FOR _bitIdx := 0 TO 15 DO
    IF (_reg.managedBitMask AND SHL(WORD#1, _bitIdx)) <> 0 THEN
        _sigIdx := _reg.arrSignalIndex[_bitIdx];

        IF _sigIdx > 0 THEN
            _pData := inpPtrWriteData + UINT_TO_DWORD(_sigIdx - 1) * SIZEOF(ST_MBWriteData);

            IF _pData^.valueBool THEN
                _baseValue := _baseValue OR SHL(WORD#1, _bitIdx);
            ELSE
                _baseValue := _baseValue AND NOT SHL(WORD#1, _bitIdx);
            END_IF
        END_IF
    END_IF
END_FOR

_reg.writeValue := _baseValue;
END_METHOD

METHOD PRIVATE checkReadComplete : BOOL
CASE _arrReadBlocks[_currentBlockIdx].functionCode OF
    1:
        fbMbReadCoils(bExecute := FALSE);
        checkReadComplete := NOT fbMbReadCoils.bBusy;
    2:
        fbMbReadInputs(bExecute := FALSE);
        checkReadComplete := NOT fbMbReadInputs.bBusy;
    3:
        fbMbReadRegs(bExecute := FALSE);
        checkReadComplete := NOT fbMbReadRegs.bBusy;
    4:
        fbMbReadInputRegs(bExecute := FALSE);
        checkReadComplete := NOT fbMbReadInputRegs.bBusy;
ELSE
    // RMW read path uses fbMbReadRegs unconditionally.
    fbMbReadRegs(bExecute := FALSE);
    checkReadComplete := NOT fbMbReadRegs.bBusy;
END_CASE
END_METHOD

METHOD PRIVATE checkStaleData
VAR
    _i          : UINT;
    _pResult    : POINTER TO ST_MBReadResult;
    _elapsed    : TIME;
END_VAR
_elapsed := TIME() - _lastGoodReadTime;

IF _elapsed > cfgStaleThreshold THEN
    FOR _i := 1 TO cfgReadSignalCount DO
        _pResult := inpPtrReadResults + UINT_TO_DWORD(_i - 1) * SIZEOF(ST_MBReadResult);

        IF _pResult^.quality = E_SignalQuality.Good THEN
            _pResult^.quality := E_SignalQuality.UncertainStale;
        END_IF
    END_FOR
END_IF
END_METHOD

METHOD PRIVATE checkWriteComplete : BOOL
IF _state = E_DriverState.WriteWait THEN
    IF _arrWriteBlocks[_currentBlockIdx].area = E_MBArea.Coils THEN
        fbMbWriteCoils(bExecute := FALSE);
        checkWriteComplete := NOT fbMbWriteCoils.bBusy;
    ELSE
        fbMbWriteRegs(bExecute := FALSE);
        checkWriteComplete := NOT fbMbWriteRegs.bBusy;
    END_IF
ELSE
    fbMbWriteSingleReg(bExecute := FALSE);
    checkWriteComplete := NOT fbMbWriteSingleReg.bBusy;
END_IF
END_METHOD

// Recover a Faulted (or errored) driver without toggling inpEnable: it restarts from Init on
// the next cycle() — re-parses the configuration and resumes polling. No effect while disabled.
METHOD PUBLIC cmdReset : BOOL
IF inpEnable THEN
    _state := E_DriverState.Init;
    _resetRequest := TRUE;
    cmdReset := TRUE;
END_IF
END_METHOD

METHOD PRIVATE combineWords : DWORD
VAR_INPUT
    inpWord0        : WORD;
    inpWord1        : WORD;
END_VAR
IF cfgWordOrder = E_WordOrder.BigEndian THEN
    combineWords := SHL(WORD_TO_DWORD(inpWord0), 16) OR WORD_TO_DWORD(inpWord1);
ELSE
    combineWords := SHL(WORD_TO_DWORD(inpWord1), 16) OR WORD_TO_DWORD(inpWord0);
END_IF
END_METHOD

PROPERTY PUBLIC commandDelay : TIME
GET
commandDelay := cfgCommandDelay;
END_GET
SET
IF NOT _initialized THEN
    cfgCommandDelay := commandDelay;
END_IF
END_SET
END_PROPERTY

METHOD PUBLIC cycle
VAR
    _risingEnable   : BOOL;
END_VAR
_risingEnable := inpEnable AND NOT _enablePrev;
_enablePrev := inpEnable;

IF NOT inpEnable THEN
    disable();
    RETURN;
END_IF

IF _initialized AND _socketConnected THEN
    stsStatus.timeSinceLastGoodRead := TIME() - _lastGoodReadTime;
    stsStatus.timeSinceLastGoodWrite := TIME() - _lastGoodWriteTime;
END_IF

CASE _state OF

    E_DriverState.Init:
        IF _risingEnable OR _resetRequest THEN
            _resetRequest := FALSE;
            reset();
            _state := E_DriverState.ParseConfig;
        END_IF

    E_DriverState.ParseConfig:
        IF parseAllConfigs() THEN
            _state := E_DriverState.OptimizeBlocks;
        ELSE
            stsError := TRUE;
            _state := E_DriverState.Error;
        END_IF

    E_DriverState.OptimizeBlocks:
        optimizeReadBlocks();
        optimizeWriteBlocks();
        identifyBitRegisters();

        stsStatus.readBlockCount := _readBlockCount;
        stsStatus.writeBlockCount := _writeBlockCount;
        stsStatus.bitRegisterCount := _bitRegisterCount;

        _initialized := TRUE;
        _state := E_DriverState.Connecting;

    E_DriverState.Connecting:
        // Tc2_ModbusCaller manages TCP internally per FB call; no explicit connect.
        // Treat the driver as "ready to talk" once configs are parsed.
        _socketConnected := TRUE;
        _connectAttempts := 0;
        stsStatus.connected := TRUE;
        stsStatus.reconnectAttempts := 0;
        _lastGoodReadTime := TIME();
        _lastGoodWriteTime := TIME();
        _state := E_DriverState.Ready;

    E_DriverState.ConnectWait:
        // Vestigial state retained for E_DriverState compatibility; transition to Ready.
        _state := E_DriverState.Ready;

    E_DriverState.ReconnectWait:
        tonReconnectDelay(IN := TRUE, PT := cfgReconnectDelay);
        IF tonReconnectDelay.Q THEN
            tonReconnectDelay(IN := FALSE);
            _socketConnected := TRUE;
            stsStatus.connected := TRUE;
            _state := E_DriverState.Ready;
        END_IF

    E_DriverState.Disconnecting:
        // No socket to disconnect (Tc2_ModbusCaller is per-call).
        _socketConnected := FALSE;
        stsStatus.connected := FALSE;
        stsStatus.readCycleActive := FALSE;
        stsStatus.writeCycleActive := FALSE;
        _consecFailures := 0;           // the retry gets its own maxConsecFails budget
        _state := E_DriverState.DisconnectWait;

    E_DriverState.DisconnectWait:
        IF _disconnectPending THEN
            _disconnectPending := FALSE;
            tonReconnectDelay(IN := FALSE);
            _state := E_DriverState.ReconnectWait;
        ELSE
            _state := E_DriverState.Init;
        END_IF

    E_DriverState.Ready:
        tonPollInterval(IN := TRUE, PT := cfgPollInterval);
        IF tonPollInterval.Q THEN
            tonPollInterval(IN := FALSE);
            IF _readBlockCount > 0 THEN
                _state := E_DriverState.ReadStart;
                RETURN;
            END_IF
        END_IF

        tonWriteInterval(IN := TRUE, PT := cfgWriteCycleInterval);
        IF tonWriteInterval.Q THEN
            tonWriteInterval(IN := FALSE);
            IF NOT inpHoldWrites AND (_writeBlockCount > 0 OR _bitRegisterCount > 0) THEN
                _state := E_DriverState.WriteStart;
                RETURN;
            END_IF
        END_IF

        checkStaleData();

    E_DriverState.ReadStart:
        _currentBlockIdx := 1;
        _readCycleFailed := FALSE;
        stsStatus.readCycleActive := TRUE;
        _state := E_DriverState.ReadSend;

    E_DriverState.ReadSend:
        IF _currentBlockIdx > _readBlockCount THEN
            _state := E_DriverState.ReadComplete;
        ELSE
            sendReadRequest(_currentBlockIdx);
            _state := E_DriverState.ReadWait;
        END_IF

    E_DriverState.ReadWait:
        tonTimeout(IN := TRUE, PT := cfgTimeout);

        IF checkReadComplete() THEN
            tonTimeout(IN := FALSE);
            IF readSucceeded() THEN
                processReadBlock(_currentBlockIdx);
                _consecFailures := 0;
            ELSE
                handleBlockError(_currentBlockIdx, TRUE);
            END_IF
            IF _state = E_DriverState.ReadWait THEN   // the error handler may have moved us to Disconnecting/Faulted
                _state := E_DriverState.ReadDelay;
            END_IF

        ELSIF tonTimeout.Q THEN
            tonTimeout(IN := FALSE);
            handleBlockError(_currentBlockIdx, TRUE);
            IF _state = E_DriverState.ReadWait THEN   // the error handler may have moved us to Disconnecting/Faulted
                _state := E_DriverState.ReadDelay;
            END_IF
        END_IF

    E_DriverState.ReadDelay:
        tonCommandDelay(IN := TRUE, PT := cfgCommandDelay);
        IF tonCommandDelay.Q THEN
            tonCommandDelay(IN := FALSE);
            _currentBlockIdx := _currentBlockIdx + 1;
            _state := E_DriverState.ReadSend;
        END_IF

    E_DriverState.ReadComplete:
        stsStatus.readCycleActive := FALSE;
        stsStatus.totalReadCycles := stsStatus.totalReadCycles + 1;
        // Only a cycle in which EVERY block succeeded is a good read. Stamping it regardless
        // kept timeSinceLastGoodRead near zero (and stale marking off) while every read failed.
        IF NOT _readCycleFailed THEN
            _lastGoodReadTime := TIME();
            _connectAttempts := 0;      // link proven again: the reconnect budget starts over
            stsStatus.reconnectAttempts := 0;
        END_IF
        _state := E_DriverState.Ready;

    E_DriverState.WriteStart:
        _currentBlockIdx := 1;
        _writeCycleFailed := FALSE;
        _currentRmwIdx := 0;
        stsStatus.writeCycleActive := TRUE;
        _state := E_DriverState.WriteSend;

    E_DriverState.WriteSend:
        WHILE _currentBlockIdx <= _writeBlockCount DO
            IF NOT _arrWriteBlocks[_currentBlockIdx].containsBitSignals THEN
                packAndSendWriteBlock(_currentBlockIdx);
                _state := E_DriverState.WriteWait;
                RETURN;
            END_IF
            _currentBlockIdx := _currentBlockIdx + 1;
        END_WHILE

        IF _currentRmwIdx < _bitRegisterCount THEN
            _currentRmwIdx := _currentRmwIdx + 1;
            _state := E_DriverState.RmwReadSend;
        ELSE
            _state := E_DriverState.WriteComplete;
        END_IF

    E_DriverState.WriteWait:
        tonTimeout(IN := TRUE, PT := cfgTimeout);

        IF checkWriteComplete() THEN
            tonTimeout(IN := FALSE);
            IF writeSucceeded() THEN
                updateWriteStatus(_currentBlockIdx, TRUE);
                _consecFailures := 0;
            ELSE
                handleBlockError(_currentBlockIdx, FALSE);
                updateWriteStatus(_currentBlockIdx, FALSE);
            END_IF
            IF _state = E_DriverState.WriteWait THEN   // the error handler may have moved us to Disconnecting/Faulted
                _state := E_DriverState.WriteDelay;
            END_IF

        ELSIF tonTimeout.Q THEN
            tonTimeout(IN := FALSE);
            handleBlockError(_currentBlockIdx, FALSE);
            updateWriteStatus(_currentBlockIdx, FALSE);
            IF _state = E_DriverState.WriteWait THEN   // the error handler may have moved us to Disconnecting/Faulted
                _state := E_DriverState.WriteDelay;
            END_IF
        END_IF

    E_DriverState.WriteDelay:
        tonCommandDelay(IN := TRUE, PT := cfgCommandDelay);
        IF tonCommandDelay.Q THEN
            tonCommandDelay(IN := FALSE);
            _currentBlockIdx := _currentBlockIdx + 1;
            _state := E_DriverState.WriteSend;
        END_IF

    E_DriverState.RmwReadSend:
        sendRmwReadRequest(_currentRmwIdx);
        _state := E_DriverState.RmwReadWait;

    E_DriverState.RmwReadWait:
        tonTimeout(IN := TRUE, PT := cfgTimeout);

        IF checkReadComplete() THEN
            tonTimeout(IN := FALSE);
            IF readSucceeded() THEN
                _arrBitRegisters[_currentRmwIdx].readValue := _arrRawReadBuffer[0];
                _state := E_DriverState.RmwModify;
            ELSE
                handleRmwError(_currentRmwIdx);
                IF _state = E_DriverState.RmwReadWait THEN   // the error handler may have moved us to Disconnecting/Faulted
                    _state := E_DriverState.RmwDelay;
                END_IF
            END_IF

        ELSIF tonTimeout.Q THEN
            tonTimeout(IN := FALSE);
            handleRmwError(_currentRmwIdx);
            IF _state = E_DriverState.RmwReadWait THEN   // the error handler may have moved us to Disconnecting/Faulted
                _state := E_DriverState.RmwDelay;
            END_IF
        END_IF

    E_DriverState.RmwModify:
        applyBitModifications(_currentRmwIdx);
        _state := E_DriverState.RmwWriteSend;

    E_DriverState.RmwWriteSend:
        sendRmwWriteRequest(_currentRmwIdx);
        _state := E_DriverState.RmwWriteWait;

    E_DriverState.RmwWriteWait:
        tonTimeout(IN := TRUE, PT := cfgTimeout);

        IF checkWriteComplete() THEN
            tonTimeout(IN := FALSE);
            IF writeSucceeded() THEN
                updateRmwStatus(_currentRmwIdx, TRUE);
                _consecFailures := 0;
            ELSE
                handleRmwError(_currentRmwIdx);
                updateRmwStatus(_currentRmwIdx, FALSE);
            END_IF
            IF _state = E_DriverState.RmwWriteWait THEN   // the error handler may have moved us to Disconnecting/Faulted
                _state := E_DriverState.RmwDelay;
            END_IF

        ELSIF tonTimeout.Q THEN
            tonTimeout(IN := FALSE);
            handleRmwError(_currentRmwIdx);
            updateRmwStatus(_currentRmwIdx, FALSE);
            IF _state = E_DriverState.RmwWriteWait THEN   // the error handler may have moved us to Disconnecting/Faulted
                _state := E_DriverState.RmwDelay;
            END_IF
        END_IF

    E_DriverState.RmwDelay:
        tonCommandDelay(IN := TRUE, PT := cfgCommandDelay);
        IF tonCommandDelay.Q THEN
            tonCommandDelay(IN := FALSE);
            IF _currentRmwIdx < _bitRegisterCount THEN
                _currentRmwIdx := _currentRmwIdx + 1;
                _state := E_DriverState.RmwReadSend;
            ELSE
                _state := E_DriverState.WriteComplete;
            END_IF
        END_IF

    E_DriverState.WriteComplete:
        stsStatus.writeCycleActive := FALSE;
        stsStatus.totalWriteCycles := stsStatus.totalWriteCycles + 1;
        IF NOT _writeCycleFailed THEN
            _lastGoodWriteTime := TIME();
        END_IF
        _state := E_DriverState.Ready;

    E_DriverState.Error:
        stsError := TRUE;
        stsStatus.totalErrors := stsStatus.totalErrors + 1;
        _disconnectPending := TRUE;
        _state := E_DriverState.Disconnecting;

    E_DriverState.Faulted:
        stsStatus.faulted := TRUE;
        stsError := TRUE;

END_CASE

stsStatus.currentState := _state;
stsStatus.consecutiveFailures := _consecFailures;
END_METHOD

METHOD PRIVATE dintToWords
VAR_INPUT
    inpValue        : DINT;
END_VAR
VAR_OUTPUT
    stsWord0        : WORD;
    stsWord1        : WORD;
END_VAR
VAR
    _dword          : DWORD;
    _w0, _w1        : WORD;
END_VAR
_dword := DINT_TO_DWORD(inpValue);
splitDword(inpValue := _dword, stsWord0 => _w0, stsWord1 => _w1);
stsWord0 := swapBytes(_w0);
stsWord1 := swapBytes(_w1);
END_METHOD

METHOD PRIVATE disable
// Tc2_ModbusCaller has no socket to tear down explicitly.
_socketConnected := FALSE;

tonPollInterval(IN := FALSE);
tonWriteInterval(IN := FALSE);
tonCommandDelay(IN := FALSE);
tonTimeout(IN := FALSE);
tonReconnectDelay(IN := FALSE);

// Back to Init from ANY state, Faulted included: re-enabling restarts the driver. (Faulted used
// to survive a disable, which left a faulted driver dead until the PLC restarted.)
_state := E_DriverState.Init;
_resetRequest := FALSE;

_initialized := FALSE;
stsStatus.connected := FALSE;
stsStatus.readCycleActive := FALSE;
stsStatus.writeCycleActive := FALSE;
END_METHOD

METHOD PRIVATE handleBlockError
VAR_INPUT
    inpBlockIdx : UINT;
    inpIsRead   : BOOL;
END_VAR
VAR
    _block      : REFERENCE TO ST_ReadBlock;
    _i          : UINT;
    _sigIdx     : UINT;
    _pResult    : POINTER TO ST_MBReadResult;
END_VAR
_consecFailures := _consecFailures + 1;
stsStatus.totalErrors := stsStatus.totalErrors + 1;
IF inpIsRead THEN
    _readCycleFailed := TRUE;
ELSE
    _writeCycleFailed := TRUE;
END_IF

IF inpIsRead THEN
    _block REF= _arrReadBlocks[inpBlockIdx];

    FOR _i := 1 TO _block.signalCount DO
        _sigIdx := _block.arrSignalIndex[_i];
        _pResult := inpPtrReadResults + UINT_TO_DWORD(_sigIdx - 1) * SIZEOF(ST_MBReadResult);
        _pResult^.quality := E_SignalQuality.BadComm;
    END_FOR
END_IF

IF _consecFailures >= cfgMaxConsecFails THEN
    _connectAttempts := _connectAttempts + 1;
    stsStatus.reconnectAttempts := _connectAttempts;

    IF _connectAttempts >= cfgMaxReconnectAttempts THEN
        _state := E_DriverState.Faulted;
    ELSE
        _disconnectPending := TRUE;
        _state := E_DriverState.Disconnecting;
    END_IF
END_IF
END_METHOD

METHOD PRIVATE handleRmwError
VAR_INPUT
    inpRmwIdx : UINT;
END_VAR
_consecFailures := _consecFailures + 1;
stsStatus.totalErrors := stsStatus.totalErrors + 1;
_writeCycleFailed := TRUE;      // RMW runs inside the write cycle

IF _consecFailures >= cfgMaxConsecFails THEN
    _connectAttempts := _connectAttempts + 1;
    stsStatus.reconnectAttempts := _connectAttempts;

    IF _connectAttempts >= cfgMaxReconnectAttempts THEN
        _state := E_DriverState.Faulted;
    ELSE
        _disconnectPending := TRUE;
        _state := E_DriverState.Disconnecting;
    END_IF
END_IF
END_METHOD

METHOD PRIVATE identifyBitRegisters
VAR
    _i, _j          : UINT;
    _addr           : UINT;
    _bitIdx         : BYTE;
    _found          : BOOL;
END_VAR
_bitRegisterCount := 0;

FOR _i := 1 TO cfgWriteSignalCount DO
    IF _arrParsedWrite[_i].valid AND _arrParsedWrite[_i].isBitInRegister THEN
        _addr := _arrParsedWrite[_i].baseAddress;
        _bitIdx := _arrParsedWrite[_i].bitIndex;

        _found := FALSE;
        FOR _j := 1 TO _bitRegisterCount DO
            IF _arrBitRegisters[_j].address = _addr THEN
                _arrBitRegisters[_j].managedBitMask :=
                    _arrBitRegisters[_j].managedBitMask OR SHL(WORD#1, _bitIdx);
                _arrBitRegisters[_j].arrSignalIndex[_bitIdx] := _i;
                _found := TRUE;
                EXIT;
            END_IF
        END_FOR

        IF NOT _found AND _bitRegisterCount < MAX_BIT_REGISTERS THEN
            _bitRegisterCount := _bitRegisterCount + 1;
            _arrBitRegisters[_bitRegisterCount].address := _addr;
            _arrBitRegisters[_bitRegisterCount].managedBitMask := SHL(WORD#1, _bitIdx);
            _arrBitRegisters[_bitRegisterCount].arrSignalIndex[_bitIdx] := _i;
        END_IF
    END_IF
END_FOR
END_METHOD

PROPERTY PUBLIC ipAddress : STRING(15)
GET
ipAddress := cfgIpAddress;
END_GET
SET
IF NOT _initialized THEN
    cfgIpAddress := ipAddress;
END_IF
END_SET
END_PROPERTY

PROPERTY PUBLIC isReady : BOOL
GET
isReady := (_state = E_DriverState.Ready) AND _socketConnected;
END_GET
END_PROPERTY

PROPERTY PUBLIC maxConsecFails : UINT
GET
maxConsecFails := cfgMaxConsecFails;
END_GET
SET
IF NOT _initialized THEN
    cfgMaxConsecFails := MAX(1, maxConsecFails);
END_IF
END_SET
END_PROPERTY

PROPERTY PUBLIC maxReconnectAttempts : UINT
GET
maxReconnectAttempts := cfgMaxReconnectAttempts;
END_GET
SET
IF NOT _initialized THEN
    cfgMaxReconnectAttempts := maxReconnectAttempts;
END_IF
END_SET
END_PROPERTY

METHOD PRIVATE optimizeReadBlocks
VAR
    _i, _j          : UINT;
    _sortCount      : UINT;
    _currentBlock   : UINT;
    _blockStart     : UINT;
    _blockEnd       : UINT;
    _blockArea      : E_MBArea;
    _gapTolerance   : UINT;
    _maxPerBlock    : UINT;
    _nextAddr       : UINT;
    _nextEnd        : UINT;
    _temp           : UINT;
END_VAR
_sortCount := 0;
FOR _i := 1 TO cfgReadSignalCount DO
    IF _arrParsedRead[_i].valid THEN
        _sortCount := _sortCount + 1;
        _arrSortIdx[_sortCount] := _i;
    END_IF
END_FOR

IF _sortCount = 0 THEN
    _readBlockCount := 0;
    RETURN;
END_IF

FOR _i := 1 TO _sortCount - 1 DO
    FOR _j := _i + 1 TO _sortCount DO
        IF shouldSwapForSort(_arrSortIdx[_i], _arrSortIdx[_j], TRUE) THEN
            _temp := _arrSortIdx[_i];
            _arrSortIdx[_i] := _arrSortIdx[_j];
            _arrSortIdx[_j] := _temp;
        END_IF
    END_FOR
END_FOR

_currentBlock := 0;
_i := 1;

WHILE _i <= _sortCount DO
    _currentBlock := _currentBlock + 1;
    IF _currentBlock > MAX_READ_BLOCKS THEN
        _currentBlock := _currentBlock - 1;
        EXIT;
    END_IF

    _blockArea := _arrParsedRead[_arrSortIdx[_i]].area;
    _blockStart := _arrParsedRead[_arrSortIdx[_i]].baseAddress;
    _blockEnd := _blockStart + _arrParsedRead[_arrSortIdx[_i]].registerCount - 1;

    IF _blockArea = E_MBArea.Coils OR _blockArea = E_MBArea.DiscreteInputs THEN
        _gapTolerance := GAP_TOLERANCE_COILS;
        _maxPerBlock := MAX_COILS_PER_BLOCK;
    ELSE
        _gapTolerance := GAP_TOLERANCE_REGS;
        _maxPerBlock := MAX_REGS_PER_BLOCK;
    END_IF

    _arrReadBlocks[_currentBlock].area := _blockArea;
    _arrReadBlocks[_currentBlock].startAddress := _blockStart;
    _arrReadBlocks[_currentBlock].signalCount := 1;
    _arrReadBlocks[_currentBlock].arrSignalIndex[1] := _arrSortIdx[_i];
    _arrReadBlocks[_currentBlock].arrOffsetInBlock[1] := 0;
    _arrReadBlocks[_currentBlock].enabled := TRUE;

    CASE _blockArea OF
        E_MBArea.Coils:
            _arrReadBlocks[_currentBlock].functionCode := 1;
        E_MBArea.DiscreteInputs:
            _arrReadBlocks[_currentBlock].functionCode := 2;
        E_MBArea.HoldingRegisters:
            _arrReadBlocks[_currentBlock].functionCode := 3;
        E_MBArea.InputRegisters:
            _arrReadBlocks[_currentBlock].functionCode := 4;
    END_CASE

    _j := _i + 1;
    WHILE _j <= _sortCount DO
        IF _arrParsedRead[_arrSortIdx[_j]].area <> _blockArea THEN
            EXIT;
        END_IF

        _nextAddr := _arrParsedRead[_arrSortIdx[_j]].baseAddress;
        _nextEnd := _nextAddr + _arrParsedRead[_arrSortIdx[_j]].registerCount - 1;

        IF _nextAddr > (_blockEnd + _gapTolerance + 1) THEN
            EXIT;
        END_IF

        IF (_nextEnd - _blockStart + 1) > _maxPerBlock THEN
            EXIT;
        END_IF

        _arrReadBlocks[_currentBlock].signalCount :=
            _arrReadBlocks[_currentBlock].signalCount + 1;
        _arrReadBlocks[_currentBlock].arrSignalIndex[_arrReadBlocks[_currentBlock].signalCount] :=
            _arrSortIdx[_j];
        _arrReadBlocks[_currentBlock].arrOffsetInBlock[_arrReadBlocks[_currentBlock].signalCount] :=
            _nextAddr - _blockStart;

        IF _nextEnd > _blockEnd THEN
            _blockEnd := _nextEnd;
        END_IF

        _j := _j + 1;
    END_WHILE

    _arrReadBlocks[_currentBlock].quantity := _blockEnd - _blockStart + 1;
    _i := _j;
END_WHILE

_readBlockCount := _currentBlock;
END_METHOD

METHOD PRIVATE optimizeWriteBlocks
VAR
    _i, _j          : UINT;
    _sortCount      : UINT;
    _currentBlock   : UINT;
    _blockStart     : UINT;
    _blockEnd       : UINT;
    _blockArea      : E_MBArea;
    _gapTolerance   : UINT;
    _maxPerBlock    : UINT;
    _nextAddr       : UINT;
    _nextEnd        : UINT;
    _temp           : UINT;
END_VAR
_sortCount := 0;
FOR _i := 1 TO cfgWriteSignalCount DO
    IF _arrParsedWrite[_i].valid AND NOT _arrParsedWrite[_i].isBitInRegister THEN
        _sortCount := _sortCount + 1;
        _arrSortIdx[_sortCount] := _i;
    END_IF
END_FOR

IF _sortCount = 0 THEN
    _writeBlockCount := 0;
    RETURN;
END_IF

FOR _i := 1 TO _sortCount - 1 DO
    FOR _j := _i + 1 TO _sortCount DO
        IF shouldSwapForSort(_arrSortIdx[_i], _arrSortIdx[_j], FALSE) THEN
            _temp := _arrSortIdx[_i];
            _arrSortIdx[_i] := _arrSortIdx[_j];
            _arrSortIdx[_j] := _temp;
        END_IF
    END_FOR
END_FOR

_currentBlock := 0;
_i := 1;

WHILE _i <= _sortCount DO
    _currentBlock := _currentBlock + 1;
    IF _currentBlock > MAX_WRITE_BLOCKS THEN
        _currentBlock := _currentBlock - 1;
        EXIT;
    END_IF

    _blockArea := _arrParsedWrite[_arrSortIdx[_i]].area;
    _blockStart := _arrParsedWrite[_arrSortIdx[_i]].baseAddress;
    _blockEnd := _blockStart + _arrParsedWrite[_arrSortIdx[_i]].registerCount - 1;

    IF _blockArea = E_MBArea.Coils THEN
        _gapTolerance := GAP_TOLERANCE_COILS;
        _maxPerBlock := MAX_COILS_PER_BLOCK;
    ELSE
        _gapTolerance := GAP_TOLERANCE_REGS;
        _maxPerBlock := MAX_REGS_PER_BLOCK;
    END_IF

    _arrWriteBlocks[_currentBlock].area := _blockArea;
    _arrWriteBlocks[_currentBlock].startAddress := _blockStart;
    _arrWriteBlocks[_currentBlock].signalCount := 1;
    _arrWriteBlocks[_currentBlock].arrSignalIndex[1] := _arrSortIdx[_i];
    _arrWriteBlocks[_currentBlock].arrOffsetInBlock[1] := 0;
    _arrWriteBlocks[_currentBlock].enabled := TRUE;
    _arrWriteBlocks[_currentBlock].containsBitSignals := FALSE;

    CASE _blockArea OF
        E_MBArea.Coils:
            _arrWriteBlocks[_currentBlock].functionCode := 15;
        E_MBArea.HoldingRegisters:
            _arrWriteBlocks[_currentBlock].functionCode := 16;
    END_CASE

    _j := _i + 1;
    WHILE _j <= _sortCount DO
        IF _arrParsedWrite[_arrSortIdx[_j]].area <> _blockArea THEN
            EXIT;
        END_IF

        _nextAddr := _arrParsedWrite[_arrSortIdx[_j]].baseAddress;
        _nextEnd := _nextAddr + _arrParsedWrite[_arrSortIdx[_j]].registerCount - 1;

        IF _nextAddr > (_blockEnd + _gapTolerance + 1) THEN
            EXIT;
        END_IF

        IF (_nextEnd - _blockStart + 1) > _maxPerBlock THEN
            EXIT;
        END_IF

        _arrWriteBlocks[_currentBlock].signalCount :=
            _arrWriteBlocks[_currentBlock].signalCount + 1;
        _arrWriteBlocks[_currentBlock].arrSignalIndex[_arrWriteBlocks[_currentBlock].signalCount] :=
            _arrSortIdx[_j];
        _arrWriteBlocks[_currentBlock].arrOffsetInBlock[_arrWriteBlocks[_currentBlock].signalCount] :=
            _nextAddr - _blockStart;

        IF _nextEnd > _blockEnd THEN
            _blockEnd := _nextEnd;
        END_IF

        _j := _j + 1;
    END_WHILE

    _arrWriteBlocks[_currentBlock].quantity := _blockEnd - _blockStart + 1;
    _i := _j;
END_WHILE

_writeBlockCount := _currentBlock;
END_METHOD

METHOD PRIVATE packAndSendWriteBlock
VAR_INPUT
    inpBlockIdx : UINT;
END_VAR
VAR
    _block      : REFERENCE TO ST_WriteBlock;
    _i          : UINT;
    _sigIdx     : UINT;
    _offset     : UINT;
    _parsed     : REFERENCE TO ST_ParsedSignal;
    _pData      : POINTER TO ST_MBWriteData;
END_VAR
_block REF= _arrWriteBlocks[inpBlockIdx];

MEMSET(ADR(_arrRawWriteBuffer), 0, SIZEOF(_arrRawWriteBuffer));

FOR _i := 1 TO _block.signalCount DO
    _sigIdx := _block.arrSignalIndex[_i];
    _offset := _block.arrOffsetInBlock[_i];
    _parsed REF= _arrParsedWrite[_sigIdx];

    _pData := inpPtrWriteData + UINT_TO_DWORD(_sigIdx - 1) * SIZEOF(ST_MBWriteData);

    CASE _parsed.dataType OF
        E_MBDataType.mbReal32:
            realToWords(
                inpValue := _pData^.valueReal,
                stsWord0 => _arrRawWriteBuffer[_offset],
                stsWord1 => _arrRawWriteBuffer[_offset + 1]
            );

        E_MBDataType.mbInt32:
            dintToWords(
                inpValue := _pData^.valueDint,
                stsWord0 => _arrRawWriteBuffer[_offset],
                stsWord1 => _arrRawWriteBuffer[_offset + 1]
            );

        E_MBDataType.mbUInt32:
            udintToWords(
                inpValue := _pData^.valueUdint,
                stsWord0 => _arrRawWriteBuffer[_offset],
                stsWord1 => _arrRawWriteBuffer[_offset + 1]
            );

        E_MBDataType.mbInt16:
            _arrRawWriteBuffer[_offset] := swapBytes(INT_TO_WORD(_pData^.valueInt));

        E_MBDataType.mbUInt16:
            _arrRawWriteBuffer[_offset] := swapBytes(UINT_TO_WORD(_pData^.valueUint));

        E_MBDataType.mbWord16:
            _arrRawWriteBuffer[_offset] := swapBytes(_pData^.valueWord);

        E_MBDataType.mbBit:
            IF _pData^.valueBool THEN
                _arrRawWriteBuffer[_offset / 16] :=
                    _arrRawWriteBuffer[_offset / 16] OR SHL(WORD#1, _offset MOD 16);
            END_IF
    END_CASE
END_FOR

IF _block.area = E_MBArea.Coils THEN
    fbMbWriteCoils(
        sIPAddr     := cfgIpAddress,
        nTCPPort    := cfgPort,
        nUnitID     := cfgUnitId,
        nQuantity   := _block.quantity,
        nMBAddr     := _block.startAddress,
        cbLength    := UINT_TO_UDINT(_block.quantity + 7) / 8,
        pSrcAddr    := ADR(_arrRawWriteBuffer),
        bExecute    := TRUE,
        tTimeout    := cfgTimeout
    );
ELSE
    fbMbWriteRegs(
        sIPAddr     := cfgIpAddress,
        nTCPPort    := cfgPort,
        nUnitID     := cfgUnitId,
        nQuantity   := _block.quantity,
        nMBAddr     := _block.startAddress,
        cbLength    := UINT_TO_UDINT(_block.quantity) * 2,
        pSrcAddr    := ADR(_arrRawWriteBuffer),
        bExecute    := TRUE,
        tTimeout    := cfgTimeout
    );
END_IF
END_METHOD

METHOD PRIVATE parseAllConfigs : BOOL
VAR
    _i              : UINT;
    _pConfig        : POINTER TO ST_MBSignalConfig;
    _pResult        : POINTER TO ST_MBReadResult;
END_VAR
IF cfgReadSignalCount > 0 AND (inpPtrReadConfig = 0 OR inpPtrReadResults = 0) THEN
    stsErrorId := 16#8001;
    RETURN;
END_IF

IF cfgWriteSignalCount > 0 AND (inpPtrWriteConfig = 0 OR inpPtrWriteData = 0) THEN
    stsErrorId := 16#8002;
    RETURN;
END_IF

FOR _i := 1 TO cfgReadSignalCount DO
    _pConfig := inpPtrReadConfig + UINT_TO_DWORD(_i - 1) * SIZEOF(ST_MBSignalConfig);

    parseModbusAddress(
        inpModbusAddr := _pConfig^.modbusAddr,
        inpDataType := _pConfig^.dataType,
        inpBitIndex := _pConfig^.bitIndex,
        stsParsed => _arrParsedRead[_i]
    );

    IF NOT _arrParsedRead[_i].valid THEN
        _pResult := inpPtrReadResults + UINT_TO_DWORD(_i - 1) * SIZEOF(ST_MBReadResult);
        _pResult^.quality := E_SignalQuality.BadConfig;
    END_IF
END_FOR

FOR _i := 1 TO cfgWriteSignalCount DO
    _pConfig := inpPtrWriteConfig + UINT_TO_DWORD(_i - 1) * SIZEOF(ST_MBSignalConfig);

    parseModbusAddress(
        inpModbusAddr := _pConfig^.modbusAddr,
        inpDataType := _pConfig^.dataType,
        inpBitIndex := _pConfig^.bitIndex,
        stsParsed => _arrParsedWrite[_i]
    );
END_FOR

parseAllConfigs := TRUE;
END_METHOD

METHOD PRIVATE parseModbusAddress
VAR_INPUT
    inpModbusAddr   : UDINT;
    inpDataType     : E_MBDataType;
    inpBitIndex     : BYTE;
END_VAR
VAR_OUTPUT
    stsParsed       : ST_ParsedSignal;
END_VAR
VAR
    _areaCode       : UDINT;
    _offset         : UDINT;
END_VAR
stsParsed.valid := FALSE;
stsParsed.dataType := inpDataType;
stsParsed.bitIndex := inpBitIndex;

IF inpModbusAddr >= 400001 THEN
    _areaCode := 4;
    _offset := (inpModbusAddr MOD 100000) - 1;
ELSIF inpModbusAddr >= 40001 THEN
    _areaCode := 4;
    _offset := (inpModbusAddr MOD 10000) - 1;
ELSIF inpModbusAddr >= 30001 THEN
    _areaCode := 3;
    _offset := (inpModbusAddr MOD 10000) - 1;
ELSIF inpModbusAddr >= 10001 THEN
    _areaCode := 1;
    _offset := (inpModbusAddr MOD 10000) - 1;
ELSIF inpModbusAddr >= 1 THEN
    _areaCode := 0;
    _offset := inpModbusAddr - 1;
ELSE
    RETURN;
END_IF

IF _offset > 65535 THEN
    RETURN;
END_IF

stsParsed.baseAddress := UDINT_TO_UINT(_offset);

CASE _areaCode OF
    0:
        stsParsed.area := E_MBArea.Coils;
        stsParsed.registerCount := 1;
        stsParsed.bitIndex := BIT_INDEX_NA;
        stsParsed.isBitInRegister := FALSE;

    1:
        stsParsed.area := E_MBArea.DiscreteInputs;
        stsParsed.registerCount := 1;
        stsParsed.bitIndex := BIT_INDEX_NA;
        stsParsed.isBitInRegister := FALSE;

    3:
        stsParsed.area := E_MBArea.InputRegisters;
        IF inpDataType = E_MBDataType.mbBit AND inpBitIndex < 16 THEN
            stsParsed.isBitInRegister := TRUE;
        END_IF

    4:
        stsParsed.area := E_MBArea.HoldingRegisters;
        IF inpDataType = E_MBDataType.mbBit AND inpBitIndex < 16 THEN
            stsParsed.isBitInRegister := TRUE;
        END_IF

ELSE
    RETURN;
END_CASE

CASE inpDataType OF
    E_MBDataType.mbReal32,
    E_MBDataType.mbInt32,
    E_MBDataType.mbUInt32:
        stsParsed.registerCount := 2;

    E_MBDataType.mbInt16,
    E_MBDataType.mbUInt16,
    E_MBDataType.mbWord16,
    E_MBDataType.mbBit:
        stsParsed.registerCount := 1;
END_CASE

stsParsed.valid := TRUE;
END_METHOD

PROPERTY PUBLIC pollInterval : TIME
GET
pollInterval := cfgPollInterval;
END_GET
SET
IF NOT _initialized THEN
    cfgPollInterval := pollInterval;
END_IF
END_SET
END_PROPERTY

PROPERTY PUBLIC port : UINT
GET
port := cfgPort;
END_GET
SET
IF NOT _initialized THEN
    cfgPort := port;
END_IF
END_SET
END_PROPERTY

METHOD PRIVATE processReadBlock
VAR_INPUT
    inpBlockIdx : UINT;
END_VAR
VAR
    _block      : REFERENCE TO ST_ReadBlock;
    _i          : UINT;
    _sigIdx     : UINT;
    _offset     : UINT;
    _parsed     : REFERENCE TO ST_ParsedSignal;
    _pResult    : POINTER TO ST_MBReadResult;
    _rawWord    : WORD;
END_VAR
_block REF= _arrReadBlocks[inpBlockIdx];

FOR _i := 1 TO _block.signalCount DO
    _sigIdx := _block.arrSignalIndex[_i];
    _offset := _block.arrOffsetInBlock[_i];
    _parsed REF= _arrParsedRead[_sigIdx];

    _pResult := inpPtrReadResults + UINT_TO_DWORD(_sigIdx - 1) * SIZEOF(ST_MBReadResult);

    CASE _parsed.dataType OF
        E_MBDataType.mbReal32:
            _pResult^.valueReal := wordsToReal(
                _arrRawReadBuffer[_offset],
                _arrRawReadBuffer[_offset + 1]
            );

        E_MBDataType.mbInt32:
            _pResult^.valueDint := wordsToDint(
                _arrRawReadBuffer[_offset],
                _arrRawReadBuffer[_offset + 1]
            );

        E_MBDataType.mbUInt32:
            _pResult^.valueUdint := wordsToUdint(
                _arrRawReadBuffer[_offset],
                _arrRawReadBuffer[_offset + 1]
            );

        E_MBDataType.mbInt16:
            _rawWord := swapBytes(_arrRawReadBuffer[_offset]);
            _pResult^.valueInt := WORD_TO_INT(_rawWord);

        E_MBDataType.mbUInt16:
            _rawWord := swapBytes(_arrRawReadBuffer[_offset]);
            _pResult^.valueUint := WORD_TO_UINT(_rawWord);

        E_MBDataType.mbWord16:
            _pResult^.valueWord := swapBytes(_arrRawReadBuffer[_offset]);

        E_MBDataType.mbBit:
            IF _parsed.isBitInRegister THEN
                _rawWord := swapBytes(_arrRawReadBuffer[_offset]);
                _pResult^.valueBool := (_rawWord AND SHL(WORD#1, _parsed.bitIndex)) <> 0;
            ELSE
                _pResult^.valueBool := (_arrRawReadBuffer[_offset / 16] AND SHL(WORD#1, _offset MOD 16)) <> 0;
            END_IF
    END_CASE

    _pResult^.quality := E_SignalQuality.Good;
    _pResult^.updateCount := _pResult^.updateCount + 1;
END_FOR
END_METHOD

PROPERTY PUBLIC readSignalCount : UINT
GET
readSignalCount := cfgReadSignalCount;
END_GET
SET
IF NOT _initialized THEN
    cfgReadSignalCount := MIN(readSignalCount, MAX_READ_SIGNALS);
END_IF
END_SET
END_PROPERTY

METHOD PRIVATE readSucceeded : BOOL
// During an RMW read, _state = RmwReadWait and there is no current read block;
// the active FB in that case is fbMbReadRegs.
IF _state = E_DriverState.RmwReadWait THEN
    readSucceeded := NOT fbMbReadRegs.bError;
    IF fbMbReadRegs.bError THEN
        _lastMbError := 1;
    END_IF
ELSE
    CASE _arrReadBlocks[_currentBlockIdx].functionCode OF
        1:
            readSucceeded := NOT fbMbReadCoils.bError;
            IF fbMbReadCoils.bError THEN
                _lastMbError := 1;
            END_IF
        2:
            readSucceeded := NOT fbMbReadInputs.bError;
            IF fbMbReadInputs.bError THEN
                _lastMbError := 1;
            END_IF
        3:
            readSucceeded := NOT fbMbReadRegs.bError;
            IF fbMbReadRegs.bError THEN
                _lastMbError := 1;
            END_IF
        4:
            readSucceeded := NOT fbMbReadInputRegs.bError;
            IF fbMbReadInputRegs.bError THEN
                _lastMbError := 1;
            END_IF
    END_CASE
END_IF

stsStatus.lastErrorCode := _lastMbError;
END_METHOD

METHOD PRIVATE realToWords
VAR_INPUT
    inpValue        : REAL;
END_VAR
VAR_OUTPUT
    stsWord0        : WORD;
    stsWord1        : WORD;
END_VAR
VAR
    _dword          : DWORD;
    _w0, _w1        : WORD;
END_VAR
MEMCPY(ADR(_dword), ADR(inpValue), SIZEOF(REAL));
splitDword(inpValue := _dword, stsWord0 => _w0, stsWord1 => _w1);
stsWord0 := swapBytes(_w0);
stsWord1 := swapBytes(_w1);
END_METHOD

PROPERTY PUBLIC reconnectDelay : TIME
GET
reconnectDelay := cfgReconnectDelay;
END_GET
SET
IF NOT _initialized THEN
    cfgReconnectDelay := reconnectDelay;
END_IF
END_SET
END_PROPERTY

METHOD PRIVATE reset
VAR
    _i : UINT;
    _pResult : POINTER TO ST_MBReadResult;
END_VAR
_state := E_DriverState.Init;
_initialized := FALSE;
_socketConnected := FALSE;
_consecFailures := 0;
_connectAttempts := 0;
_disconnectPending := FALSE;

MEMSET(ADR(stsStatus), 0, SIZEOF(stsStatus));
stsError := FALSE;
stsErrorId := 0;

MEMSET(ADR(_arrParsedRead), 0, SIZEOF(_arrParsedRead));
MEMSET(ADR(_arrParsedWrite), 0, SIZEOF(_arrParsedWrite));
MEMSET(ADR(_arrReadBlocks), 0, SIZEOF(_arrReadBlocks));
MEMSET(ADR(_arrWriteBlocks), 0, SIZEOF(_arrWriteBlocks));
MEMSET(ADR(_arrBitRegisters), 0, SIZEOF(_arrBitRegisters));

_readBlockCount := 0;
_writeBlockCount := 0;
_bitRegisterCount := 0;

tonPollInterval(IN := FALSE);
tonWriteInterval(IN := FALSE);
tonCommandDelay(IN := FALSE);
tonTimeout(IN := FALSE);
tonReconnectDelay(IN := FALSE);

IF inpPtrReadResults <> 0 THEN
    FOR _i := 1 TO cfgReadSignalCount DO
        _pResult := inpPtrReadResults + UINT_TO_DWORD(_i - 1) * SIZEOF(ST_MBReadResult);
        _pResult^.quality := E_SignalQuality.UncertainInit;
    END_FOR
END_IF
END_METHOD

METHOD PRIVATE sendReadRequest
VAR_INPUT
    inpBlockIdx : UINT;
END_VAR
VAR
    _block : REFERENCE TO ST_ReadBlock;
END_VAR
_block REF= _arrReadBlocks[inpBlockIdx];

CASE _block.functionCode OF
    1:  // FC01 Read Coils
        fbMbReadCoils(
            sIPAddr     := cfgIpAddress,
            nTCPPort    := cfgPort,
            nUnitID     := cfgUnitId,
            nQuantity   := _block.quantity,
            nMBAddr     := _block.startAddress,
            cbLength    := SIZEOF(_arrRawReadBuffer),
            pDestAddr   := ADR(_arrRawReadBuffer),
            bExecute    := TRUE,
            tTimeout    := cfgTimeout
        );

    2:  // FC02 Read Discrete Inputs
        fbMbReadInputs(
            sIPAddr     := cfgIpAddress,
            nTCPPort    := cfgPort,
            nUnitID     := cfgUnitId,
            nQuantity   := _block.quantity,
            nMBAddr     := _block.startAddress,
            cbLength    := SIZEOF(_arrRawReadBuffer),
            pDestAddr   := ADR(_arrRawReadBuffer),
            bExecute    := TRUE,
            tTimeout    := cfgTimeout
        );

    3:  // FC03 Read Holding Registers
        fbMbReadRegs(
            sIPAddr     := cfgIpAddress,
            nTCPPort    := cfgPort,
            nUnitID     := cfgUnitId,
            nQuantity   := _block.quantity,
            nMBAddr     := _block.startAddress,
            cbLength    := UINT_TO_UDINT(_block.quantity) * 2,
            pDestAddr   := ADR(_arrRawReadBuffer),
            bExecute    := TRUE,
            tTimeout    := cfgTimeout
        );

    4:  // FC04 Read Input Registers
        fbMbReadInputRegs(
            sIPAddr     := cfgIpAddress,
            nTCPPort    := cfgPort,
            nUnitID     := cfgUnitId,
            nQuantity   := _block.quantity,
            nMBAddr     := _block.startAddress,
            cbLength    := UINT_TO_UDINT(_block.quantity) * 2,
            pDestAddr   := ADR(_arrRawReadBuffer),
            bExecute    := TRUE,
            tTimeout    := cfgTimeout
        );
END_CASE
END_METHOD

METHOD PRIVATE sendRmwReadRequest
VAR_INPUT
    inpRmwIdx : UINT;
END_VAR
// RMW always operates on a single holding register (FC03 read).
fbMbReadRegs(
    sIPAddr     := cfgIpAddress,
    nTCPPort    := cfgPort,
    nUnitID     := cfgUnitId,
    nQuantity   := 1,
    nMBAddr     := _arrBitRegisters[inpRmwIdx].address,
    cbLength    := 2,
    pDestAddr   := ADR(_arrRawReadBuffer),
    bExecute    := TRUE,
    tTimeout    := cfgTimeout
);
END_METHOD

METHOD PRIVATE sendRmwWriteRequest
VAR_INPUT
    inpRmwIdx : UINT;
END_VAR
fbMbWriteSingleReg(
    sIPAddr     := cfgIpAddress,
    nTCPPort    := cfgPort,
    nUnitID     := cfgUnitId,
    nMBAddr     := _arrBitRegisters[inpRmwIdx].address,
    nValue      := swapBytes(_arrBitRegisters[inpRmwIdx].writeValue),
    bExecute    := TRUE,
    tTimeout    := cfgTimeout
);
END_METHOD

METHOD PRIVATE shouldSwapForSort : BOOL
VAR_INPUT
    inpIdx1         : UINT;
    inpIdx2         : UINT;
    inpIsRead       : BOOL;
END_VAR
VAR
    _area1, _area2  : E_MBArea;
    _addr1, _addr2  : UINT;
END_VAR
IF inpIsRead THEN
    _area1 := _arrParsedRead[inpIdx1].area;
    _area2 := _arrParsedRead[inpIdx2].area;
    _addr1 := _arrParsedRead[inpIdx1].baseAddress;
    _addr2 := _arrParsedRead[inpIdx2].baseAddress;
ELSE
    _area1 := _arrParsedWrite[inpIdx1].area;
    _area2 := _arrParsedWrite[inpIdx2].area;
    _addr1 := _arrParsedWrite[inpIdx1].baseAddress;
    _addr2 := _arrParsedWrite[inpIdx2].baseAddress;
END_IF

IF _area1 > _area2 THEN
    shouldSwapForSort := TRUE;
ELSIF _area1 = _area2 AND _addr1 > _addr2 THEN
    shouldSwapForSort := TRUE;
ELSE
    shouldSwapForSort := FALSE;
END_IF
END_METHOD

METHOD PRIVATE splitDword
VAR_INPUT
    inpValue        : DWORD;
END_VAR
VAR_OUTPUT
    stsWord0        : WORD;
    stsWord1        : WORD;
END_VAR
IF cfgWordOrder = E_WordOrder.BigEndian THEN
    stsWord0 := DWORD_TO_WORD(SHR(inpValue, 16));
    stsWord1 := DWORD_TO_WORD(inpValue AND 16#FFFF);
ELSE
    stsWord0 := DWORD_TO_WORD(inpValue AND 16#FFFF);
    stsWord1 := DWORD_TO_WORD(SHR(inpValue, 16));
END_IF
END_METHOD

PROPERTY PUBLIC staleThreshold : TIME
GET
staleThreshold := cfgStaleThreshold;
END_GET
SET
IF NOT _initialized THEN
    cfgStaleThreshold := staleThreshold;
END_IF
END_SET
END_PROPERTY

METHOD PRIVATE swapBytes : WORD
VAR_INPUT
    inpValue : WORD;
END_VAR
// Tc2_ModbusCaller (FB_MBReadRegs / FB_MBWriteRegs) already converts between
// network and host byte order — each WORD in _arrRawReadBuffer / _arrRawWriteBuffer
// is already the correct host-order register value. No additional byte swap needed.
swapBytes := inpValue;
END_METHOD

PROPERTY PUBLIC timeout : TIME
GET
timeout := cfgTimeout;
END_GET
SET
IF NOT _initialized THEN
    cfgTimeout := timeout;
END_IF
END_SET
END_PROPERTY

METHOD PRIVATE udintToWords
VAR_INPUT
    inpValue        : UDINT;
END_VAR
VAR_OUTPUT
    stsWord0        : WORD;
    stsWord1        : WORD;
END_VAR
VAR
    _dword          : DWORD;
    _w0, _w1        : WORD;
END_VAR
_dword := UDINT_TO_DWORD(inpValue);
splitDword(inpValue := _dword, stsWord0 => _w0, stsWord1 => _w1);
stsWord0 := swapBytes(_w0);
stsWord1 := swapBytes(_w1);
END_METHOD

PROPERTY PUBLIC unitId : BYTE
GET
unitId := cfgUnitId;
END_GET
SET
IF NOT _initialized THEN
    cfgUnitId := unitId;
END_IF
END_SET
END_PROPERTY

METHOD PRIVATE updateRmwStatus
VAR_INPUT
    inpRmwIdx   : UINT;
    inpSuccess  : BOOL;
END_VAR
VAR
    _reg        : REFERENCE TO ST_BitRegisterRmw;
    _bitIdx     : UINT;
    _sigIdx     : UINT;
    _pData      : POINTER TO ST_MBWriteData;
END_VAR
_reg REF= _arrBitRegisters[inpRmwIdx];

FOR _bitIdx := 0 TO 15 DO
    IF (_reg.managedBitMask AND SHL(WORD#1, _bitIdx)) <> 0 THEN
        _sigIdx := _reg.arrSignalIndex[_bitIdx];

        IF _sigIdx > 0 THEN
            _pData := inpPtrWriteData + UINT_TO_DWORD(_sigIdx - 1) * SIZEOF(ST_MBWriteData);

            _pData^.writeSuccess := inpSuccess;
            _pData^.writeError := NOT inpSuccess;

            IF inpSuccess THEN
                _pData^.writeCount := _pData^.writeCount + 1;
            END_IF
        END_IF
    END_IF
END_FOR
END_METHOD

METHOD PRIVATE updateWriteStatus
VAR_INPUT
    inpBlockIdx : UINT;
    inpSuccess  : BOOL;
END_VAR
VAR
    _block      : REFERENCE TO ST_WriteBlock;
    _i          : UINT;
    _sigIdx     : UINT;
    _pData      : POINTER TO ST_MBWriteData;
END_VAR
_block REF= _arrWriteBlocks[inpBlockIdx];

FOR _i := 1 TO _block.signalCount DO
    _sigIdx := _block.arrSignalIndex[_i];
    _pData := inpPtrWriteData + UINT_TO_DWORD(_sigIdx - 1) * SIZEOF(ST_MBWriteData);

    _pData^.writeSuccess := inpSuccess;
    _pData^.writeError := NOT inpSuccess;

    IF inpSuccess THEN
        _pData^.writeCount := _pData^.writeCount + 1;
    END_IF
END_FOR
END_METHOD

PROPERTY PUBLIC wordOrder : E_WordOrder
GET
wordOrder := cfgWordOrder;
END_GET
SET
IF NOT _initialized THEN
    cfgWordOrder := wordOrder;
END_IF
END_SET
END_PROPERTY

METHOD PRIVATE wordsToDint : DINT
VAR_INPUT
    inpWord0        : WORD;
    inpWord1        : WORD;
END_VAR
VAR
    _w0             : WORD;
    _w1             : WORD;
    _dword          : DWORD;
END_VAR
_w0 := swapBytes(inpWord0);
_w1 := swapBytes(inpWord1);
_dword := combineWords(_w0, _w1);
wordsToDint := DWORD_TO_DINT(_dword);
END_METHOD

METHOD PRIVATE wordsToReal : REAL
VAR_INPUT
    inpWord0        : WORD;
    inpWord1        : WORD;
END_VAR
VAR
    _w0             : WORD;
    _w1             : WORD;
    _dword          : DWORD;
    _result         : REAL;
END_VAR
_w0 := swapBytes(inpWord0);
_w1 := swapBytes(inpWord1);
_dword := combineWords(_w0, _w1);
MEMCPY(ADR(_result), ADR(_dword), SIZEOF(REAL));
wordsToReal := _result;
END_METHOD

METHOD PRIVATE wordsToUdint : UDINT
VAR_INPUT
    inpWord0        : WORD;
    inpWord1        : WORD;
END_VAR
VAR
    _w0             : WORD;
    _w1             : WORD;
    _dword          : DWORD;
END_VAR
_w0 := swapBytes(inpWord0);
_w1 := swapBytes(inpWord1);
_dword := combineWords(_w0, _w1);
wordsToUdint := DWORD_TO_UDINT(_dword);
END_METHOD

PROPERTY PUBLIC writeCycleInterval : TIME
GET
writeCycleInterval := cfgWriteCycleInterval;
END_GET
SET
IF NOT _initialized THEN
    cfgWriteCycleInterval := writeCycleInterval;
END_IF
END_SET
END_PROPERTY

PROPERTY PUBLIC writeSignalCount : UINT
GET
writeSignalCount := cfgWriteSignalCount;
END_GET
SET
IF NOT _initialized THEN
    cfgWriteSignalCount := MIN(writeSignalCount, MAX_WRITE_SIGNALS);
END_IF
END_SET
END_PROPERTY

METHOD PRIVATE writeSucceeded : BOOL
IF _state = E_DriverState.WriteWait THEN
    IF _arrWriteBlocks[_currentBlockIdx].area = E_MBArea.Coils THEN
        writeSucceeded := NOT fbMbWriteCoils.bError;
        IF fbMbWriteCoils.bError THEN
            _lastMbError := 1;
        END_IF
    ELSE
        writeSucceeded := NOT fbMbWriteRegs.bError;
        IF fbMbWriteRegs.bError THEN
            _lastMbError := 1;
        END_IF
    END_IF
ELSE
    writeSucceeded := NOT fbMbWriteSingleReg.bError;
    IF fbMbWriteSingleReg.bError THEN
        _lastMbError := 1;
    END_IF
END_IF

stsStatus.lastErrorCode := _lastMbError;
END_METHOD

END_FUNCTION_BLOCK

// ---- POUs/FBs/Comm/fb_MQTT_Connector.TcPOU
// ═══════════════════════════════════════════════════════════════════════
// fb_MQTT_Connector
// Generic MQTT signal connector with registration pattern
//
// Features:
//   - Register signals at runtime with type information
//   - Publish on change-of-state or periodic interval
//   - Transaction group publishing (multiple signals as JSON)
//   - Subscribe to topics and write values to PLC variables
//   - Bidirectional signals supported
//   - Separate publish/subscribe base topics
//   - Online change detection with automatic re-registration prompt
//   - Fault handling with configurable failure threshold
//
// Usage:
//   1. Configure cfgClientID, cfgBrokerIP, cfgPublishBaseTopic, cfgSubscribeBaseTopic
//   2. Call RegisterSignal() for each signal
//   3. Call AcknowledgeOnlineChange() after registration complete
//   4. Call Run() every scan cycle
//   5. Handle stsOnlineChangeDetected by re-registering signals
//
// ═══════════════════════════════════════════════════════════════════════
{attribute 'no_assign'}
FUNCTION_BLOCK fb_MQTT_Connector
VAR_INPUT
    // Configuration (set once at startup)
    cfgClientID             : STRING(80);       // MQTT client ID
    cfgBrokerIP             : STRING(80);       // Broker hostname or IP
    cfgPublishBaseTopic     : STRING(80);       // Base topic prefix for publishing
    cfgSubscribeBaseTopic   : STRING(80);       // Base topic prefix for subscriptions
    cfgPort                 : UINT := 1883;     // MQTT broker port
    cfgMaxConsecFails       : UINT := 10;       // Fault after N consecutive publish failures
    cfgPublishesPerScan     : UINT := 5;        // Max publishes per scan cycle
    cfgSubscribeQoS         : TcIotMqttQos := TcIotMqttQos.AtLeastOnceDelivery;
    cfgPublishQoS           : TcIotMqttQos := TcIotMqttQos.AtMostOnceDelivery;
    cfgRetainPublish        : BOOL := TRUE;     // Retain flag for published messages

    // Transaction group configuration
    cfgTxGroup1Period       : TIME := T#100MS;  // Transaction group 1 publish period
    cfgTxGroup2Period       : TIME := T#1S;     // Transaction group 2 publish period
    cfgTxGroup3Period       : TIME := T#5S;     // Transaction group 3 publish period
    cfgTxGroup1Topic        : STRING(80) := 'txgroup1'; // Transaction group 1 sub-topic
    cfgTxGroup2Topic        : STRING(80) := 'txgroup2'; // Transaction group 2 sub-topic
    cfgTxGroup3Topic        : STRING(80) := 'txgroup3'; // Transaction group 3 sub-topic

    // Commands (dynamic inputs)
    inpEnable               : BOOL;             // Enable MQTT connection
    inpReset                : BOOL;             // Reset fault (rising edge)
END_VAR

VAR_OUTPUT
    stsConnected            : BOOL;             // TRUE when connected to broker
    stsSubscribed           : BOOL;             // TRUE when subscribed to base topic
    stsFaulted              : BOOL;             // TRUE when faulted
    stsFaultCode            : UINT;             // Fault code (see constants)
    stsConsecFailures       : UINT;             // Current consecutive failure count
    stsRegisteredCount      : UINT;             // Number of registered signals
    stsRegistered           : BOOL;             // TRUE when registration complete
    stsOnlineChangeDetected : BOOL;             // TRUE when online change detected - re-register!
    stsTotalPublished       : UDINT;            // Lifetime published message count
    stsTotalReceived        : UDINT;            // Lifetime received message count
END_VAR

VAR CONSTANT
    MAX_SIGNALS             : UINT := 64;       // Maximum number of signals
    MAX_TX_PAYLOAD          : UDINT := 4095;    // Max JSON payload size for transaction groups
    FAULT_NONE              : UINT := 0;
    FAULT_CONNECTION        : UINT := 1;
    FAULT_PUBLISH           : UINT := 2;
    FAULT_POINTER_INVALID   : UINT := 3;
END_VAR

VAR
    // Signal registry
    _signals                : ARRAY[1..64] OF ST_MQTT_Signal;
    _signalCount            : UINT;

    // Publish engine state
    _publishIndex           : UINT := 1;        // Round-robin index
    _currentTime            : TIME;

    // Transaction group state
    _txGroupLastTime        : ARRAY[1..3] OF TIME;
    _txPayload              : STRING(4095);     // JSON build buffer
    _txLen                  : UDINT;            // running length of _txPayload (LEN() caps at 255)
    _txFirst                : BOOL;

    // MQTT client (FB instances - no underscore per convention)
    mqttClient              : FB_IotMqtt5Client;
    mqttMessage             : FB_IotMqtt5Message;

    // Connection state
    _mqttExecute            : BOOL;
    _subscribeTopicWildcard : STRING(255);
    _hasSubscribed          : BOOL;

    // Fault handling
    _consecFailures         : UINT;
    _resetTrig              : R_TRIG;

    // Receive buffer
    _receivedTopic          : STRING(255);
    _receivedPayload        : STRING(4095);

    // JSON parser
    fbJsonParser            : FB_JsonDomParser;
    _jsonDoc                : SJsonValue;
    _jsonRoot               : SJsonValue;
    _jsonParent             : SJsonValue;
    _jsonValue              : SJsonValue;
    _jsonParsed             : BOOL;
    _jsonValueStr           : STRING(255);

    // Working variables
    _fullTopic              : STRING(255);
    _publishPayload         : STRING(255);
    _i                      : UINT;
    _publishResult          : BOOL;
    _currentValue           : STRING(255);
END_VAR

// FB body is empty - all logic is in Run() method
// Call Run() every scan cycle after registration is complete

// ═══════════════════════════════════════════════════════════════════════
// METHOD AcknowledgeOnlineChange
// Call after re-registration is complete to clear the flag
// ═══════════════════════════════════════════════════════════════════════
METHOD PUBLIC AcknowledgeOnlineChange : BOOL
VAR_INPUT
END_VAR
stsOnlineChangeDetected := FALSE;
stsRegistered := (_signalCount > 0);

AcknowledgeOnlineChange := TRUE;
END_METHOD

// ═══════════════════════════════════════════════════════════════════════
// METHOD PRIVATE AppendToPayload
// Append a string to the _txPayload buffer using MEMCPY
// Handles strings larger than 255 chars (bypasses CONCAT limitation)
// Returns: TRUE if successful, FALSE if buffer would overflow
// ═══════════════════════════════════════════════════════════════════════
METHOD PRIVATE AppendToPayload : BOOL
VAR_INPUT
    inpStr : STRING(255);
END_VAR
VAR
    _curLen     : UDINT;
    _addLen     : UDINT;
END_VAR
// Use the tracked running length — LEN(_txPayload) caps at 255 and would truncate the group JSON.
_curLen := _txLen;
_addLen := INT_TO_UDINT(LEN(inpStr));

IF (_curLen + _addLen) > MAX_TX_PAYLOAD THEN
    AppendToPayload := FALSE;
    RETURN;
END_IF

MEMCPY(ADR(_txPayload) + _curLen, ADR(inpStr), _addLen);
// Null-terminate
MEMSET(ADR(_txPayload) + _curLen + _addLen, 0, 1);
_txLen := _curLen + _addLen;

AppendToPayload := TRUE;
END_METHOD

// ═══════════════════════════════════════════════════════════════════════
// METHOD ClearRegistration
// Clear all registered signals (call before re-registering)
// ═══════════════════════════════════════════════════════════════════════
METHOD PUBLIC ClearRegistration : BOOL
VAR_INPUT
END_VAR
MEMSET(ADR(_signals), 0, SIZEOF(_signals));
MEMSET(ADR(_txGroupLastTime), 0, SIZEOF(_txGroupLastTime));
_signalCount := 0;
stsRegisteredCount := 0;
stsRegistered := FALSE;
_publishIndex := 1;

ClearRegistration := TRUE;
END_METHOD

// ═══════════════════════════════════════════════════════════════════════
// METHOD PRIVATE ExtractJsonValue
// Extract a value from the already-parsed JSON DOM by key
// If inpJsonParentKey is non-empty, navigates to parent object first
// Returns: value as STRING(255), or empty string if key not found
// ═══════════════════════════════════════════════════════════════════════
METHOD PRIVATE ExtractJsonValue : STRING(255)
VAR_INPUT
    inpJsonKey       : STRING(255);
    inpJsonParentKey : STRING(80);
END_VAR
VAR
    _searchNode : SJsonValue;
    _targetNode : SJsonValue;
END_VAR
ExtractJsonValue := '';

// Start from the document root
_searchNode := _jsonRoot;

// If parent key specified, navigate into it first
IF LEN(inpJsonParentKey) > 0 THEN
    IF NOT fbJsonParser.HasMember(_searchNode, inpJsonParentKey) THEN
        RETURN;
    END_IF
    _searchNode := fbJsonParser.FindMember(_searchNode, inpJsonParentKey);
    IF NOT fbJsonParser.IsObject(_searchNode) THEN
        RETURN;
    END_IF
END_IF

// Find the target key
IF NOT fbJsonParser.HasMember(_searchNode, inpJsonKey) THEN
    RETURN;
END_IF
_targetNode := fbJsonParser.FindMember(_searchNode, inpJsonKey);

// Extract value based on JSON type
IF fbJsonParser.IsString(_targetNode) THEN
    ExtractJsonValue := fbJsonParser.GetString(_targetNode);
ELSIF fbJsonParser.IsNumber(_targetNode) THEN
    ExtractJsonValue := LREAL_TO_STRING(fbJsonParser.GetDouble(_targetNode));
ELSIF fbJsonParser.IsBool(_targetNode) THEN
    IF fbJsonParser.GetBool(_targetNode) THEN
        ExtractJsonValue := 'true';
    ELSE
        ExtractJsonValue := 'false';
    END_IF
ELSIF fbJsonParser.IsNull(_targetNode) THEN
    ExtractJsonValue := '';
END_IF
END_METHOD

// ═══════════════════════════════════════════════════════════════════════
// METHOD PRIVATE FindSignalByTopic
// Find signal index by matching full topic against subscribe base topic
// Returns: Signal index (1-based), or 0 if not found
// ═══════════════════════════════════════════════════════════════════════
METHOD PRIVATE FindSignalByTopic : UINT
VAR_INPUT
    inpFullTopic : STRING(255);
END_VAR
VAR
    _idx            : UINT;
    _expectedTopic  : STRING(255);
END_VAR
FindSignalByTopic := 0;

FOR _idx := 1 TO _signalCount DO
    IF _signals[_idx].bRegistered THEN
        _expectedTopic := CONCAT(CONCAT(cfgSubscribeBaseTopic, '/'), _signals[_idx].sSubTopic);

        IF _expectedTopic = inpFullTopic THEN
            FindSignalByTopic := _idx;
            RETURN;
        END_IF
    END_IF
END_FOR
END_METHOD

// ═══════════════════════════════════════════════════════════════════════
// METHOD PRIVATE IsPointerValid
// Basic validation that pointer is non-null and in valid memory range
// ═══════════════════════════════════════════════════════════════════════
METHOD PRIVATE IsPointerValid : BOOL
VAR_INPUT
    inpPCheck : PVOID;
END_VAR
// Null check + basic range check
// Valid data memory in TwinCAT typically starts above 0x10000
IsPointerValid := (inpPCheck <> 0) AND (inpPCheck > 16#10000);
END_METHOD

// ═══════════════════════════════════════════════════════════════════════
// METHOD RegisterSignal
// Add a signal to the registry
// Returns: Signal index (1-based), or 0 if registry full or invalid input
//
// For TRANSACTION_GROUP_x modes:
//   - inpPublishInterval is ignored (group period used instead)
//   - Signal's sSubTopic becomes the JSON key
//   - All signals in a group are published together as a JSON object
// ═══════════════════════════════════════════════════════════════════════
METHOD PUBLIC RegisterSignal : UINT
VAR_INPUT
    inpSubTopic         : STRING(80);           // Topic suffix (appended to base topic)
    inpPValue           : PVOID;                // ADR(yourVariable)
    inpType             : E_MQTT_SignalType;    // Data type
    inpPublishMode      : E_MQTT_PublishMode := E_MQTT_PublishMode.CHANGE_OF_STATE;
    inpDirection        : E_MQTT_Direction := E_MQTT_Direction.PUBLISH;
    inpPublishInterval  : TIME := T#1S;         // Only used for PERIODIC mode
    inpJsonKey          : STRING(255) := '';    // JSON key to extract (empty = raw payload)
    inpJsonParentKey    : STRING(80) := '';     // Parent object key (e.g. 'signals')
END_VAR
VAR
    _nextSlot : UINT;
END_VAR
// Validate inputs
IF inpPValue = 0 THEN
    RegisterSignal := 0;
    RETURN;
END_IF

IF inpType = E_MQTT_SignalType.NONE THEN
    RegisterSignal := 0;
    RETURN;
END_IF

// Check for space in registry
IF _signalCount >= MAX_SIGNALS THEN
    RegisterSignal := 0;
    RETURN;
END_IF

_nextSlot := _signalCount + 1;

// Populate signal descriptor
_signals[_nextSlot].sSubTopic        := inpSubTopic;
_signals[_nextSlot].pValue           := inpPValue;
_signals[_nextSlot].eType            := inpType;
_signals[_nextSlot].ePublishMode     := inpPublishMode;
_signals[_nextSlot].eDirection       := inpDirection;
_signals[_nextSlot].tPublishInterval := inpPublishInterval;
_signals[_nextSlot].sJsonKey         := inpJsonKey;
_signals[_nextSlot].sJsonParentKey   := inpJsonParentKey;
_signals[_nextSlot].sLastPublished   := '';
_signals[_nextSlot].tLastPublishTime := T#0S;
_signals[_nextSlot].bRegistered      := TRUE;
_signals[_nextSlot].nConsecFails     := 0;

_signalCount := _nextSlot;
stsRegisteredCount := _signalCount;

RegisterSignal := _nextSlot;
END_METHOD

// ═══════════════════════════════════════════════════════════════════════
// METHOD Run
// Call every scan cycle to process MQTT communication
// Returns: TRUE if running normally, FALSE if faulted or waiting
// ═══════════════════════════════════════════════════════════════════════
METHOD PUBLIC Run : BOOL
VAR_INPUT
END_VAR
VAR
    _publishCount   : UINT;
    _needsPublish   : BOOL;
    _signalIndex    : UINT;
    _txGroupIdx     : UINT;
    _txGroupPeriod  : TIME;
    _txGroupMode    : E_MQTT_PublishMode;
    _txHasSignals   : BOOL;
END_VAR
// ─────────────────────────────────────────────────────────────────────
// Reset handling (rising edge)
// ─────────────────────────────────────────────────────────────────────
_resetTrig(CLK := inpReset);
IF _resetTrig.Q THEN
    stsFaulted := FALSE;
    stsFaultCode := FAULT_NONE;
    _consecFailures := 0;
    stsConsecFailures := 0;
END_IF

// ─────────────────────────────────────────────────────────────────────
// Online change detection — REMOVED. It read _AppInfo.OnlineChangeCnt, a system global the CX7000
// target does not expose (compile errors C0046 '_AppInfo' not defined / C0032). Registered signals
// point at GLOBAL (GVL) variables whose addresses are stable across an online change, so automatic
// re-registration isn't needed here. If a caller ever DOES need to re-register (e.g. after moving a
// registered variable), it can call ClearRegistration() + RegisterSignal() itself; stsOnlineChange-
// Detected remains an output for API compatibility (it is simply never asserted now).
// ─────────────────────────────────────────────────────────────────────

// ─────────────────────────────────────────────────────────────────────
// If faulted, do nothing until reset
// ─────────────────────────────────────────────────────────────────────
IF stsFaulted THEN
    Run := FALSE;
    RETURN;
END_IF

// ─────────────────────────────────────────────────────────────────────
// If online change detected, wait for re-registration
// ─────────────────────────────────────────────────────────────────────
IF stsOnlineChangeDetected THEN
    Run := FALSE;
    RETURN;
END_IF

// ─────────────────────────────────────────────────────────────────────
// MQTT connection management
// ─────────────────────────────────────────────────────────────────────
mqttClient.sClientId := cfgClientID;
mqttClient.sHostName := cfgBrokerIP;
mqttClient.nHostPort := cfgPort;

_mqttExecute := inpEnable;
mqttClient.Execute(_mqttExecute);

stsConnected := mqttClient.bConnected;

IF NOT stsConnected THEN
    _hasSubscribed := FALSE;
    stsSubscribed := FALSE;
    Run := FALSE;
    RETURN;
END_IF

// ─────────────────────────────────────────────────────────────────────
// Subscribe to base topic wildcard (once after connection)
// ─────────────────────────────────────────────────────────────────────
IF NOT _hasSubscribed THEN
    _subscribeTopicWildcard := CONCAT(cfgSubscribeBaseTopic, '/#');
    _hasSubscribed := mqttClient.Subscribe(
        sTopic := _subscribeTopicWildcard,
        eQoS := cfgSubscribeQoS
    );
    stsSubscribed := _hasSubscribed;
END_IF

// ─────────────────────────────────────────────────────────────────────
// Get current time for interval checking
// ─────────────────────────────────────────────────────────────────────
_currentTime := TIME();

// ─────────────────────────────────────────────────────────────────────
// PUBLISH ENGINE - Round robin through registered signals
// Handles CHANGE_OF_STATE and PERIODIC modes
// (Transaction group signals are skipped here, handled below)
// ─────────────────────────────────────────────────────────────────────
_publishCount := 0;

WHILE _publishCount < cfgPublishesPerScan AND _signalCount > 0 DO

    // Wrap index back to start
    IF _publishIndex > _signalCount THEN
        _publishIndex := 1;
    END_IF

    _signalIndex := _publishIndex;
    _publishIndex := _publishIndex + 1;
    _publishCount := _publishCount + 1;

    // Skip if not registered
    IF NOT _signals[_signalIndex].bRegistered THEN
        CONTINUE;
    END_IF

    // Skip subscribe-only signals
    IF _signals[_signalIndex].eDirection = E_MQTT_Direction.SUBSCRIBE THEN
        CONTINUE;
    END_IF

    // Skip disabled publish mode
    IF _signals[_signalIndex].ePublishMode = E_MQTT_PublishMode.DISABLED THEN
        CONTINUE;
    END_IF

    // Skip transaction group signals (handled in TX group engine below)
    IF _signals[_signalIndex].ePublishMode = E_MQTT_PublishMode.TRANSACTION_GROUP_1
       OR _signals[_signalIndex].ePublishMode = E_MQTT_PublishMode.TRANSACTION_GROUP_2
       OR _signals[_signalIndex].ePublishMode = E_MQTT_PublishMode.TRANSACTION_GROUP_3 THEN
        CONTINUE;
    END_IF

    // Validate pointer before dereferencing
    IF NOT IsPointerValid(_signals[_signalIndex].pValue) THEN
        stsFaulted := TRUE;
        stsFaultCode := FAULT_POINTER_INVALID;
        Run := FALSE;
        RETURN;
    END_IF

    // Get current value as string
    _currentValue := ValueToString(
        inpPValue := _signals[_signalIndex].pValue,
        inpType := _signals[_signalIndex].eType
    );

    // Determine if publish is needed based on mode
    _needsPublish := FALSE;

    CASE _signals[_signalIndex].ePublishMode OF

        E_MQTT_PublishMode.CHANGE_OF_STATE:
            // Publish only when value changes
            IF _currentValue <> _signals[_signalIndex].sLastPublished THEN
                _needsPublish := TRUE;
            END_IF

        E_MQTT_PublishMode.PERIODIC:
            // Publish on change OR when interval elapsed
            IF _currentValue <> _signals[_signalIndex].sLastPublished THEN
                _needsPublish := TRUE;
            ELSIF (_currentTime - _signals[_signalIndex].tLastPublishTime) >= _signals[_signalIndex].tPublishInterval THEN
                _needsPublish := TRUE;
            END_IF

    END_CASE

    // Execute publish if needed
    IF _needsPublish THEN
        _fullTopic := CONCAT(CONCAT(cfgPublishBaseTopic, '/'), _signals[_signalIndex].sSubTopic);
        _publishPayload := _currentValue;

        _publishResult := mqttClient.Publish(
            sTopic := _fullTopic,
            pPayload := ADR(_publishPayload),
            nPayloadSize := INT_TO_UDINT(LEN(_publishPayload)),
            eQoS := cfgPublishQoS,
            bRetain := cfgRetainPublish
        );

        IF _publishResult THEN
            // Success - update state
            _signals[_signalIndex].sLastPublished := _currentValue;
            _signals[_signalIndex].tLastPublishTime := _currentTime;
            _signals[_signalIndex].nConsecFails := 0;
            _consecFailures := 0;
            stsTotalPublished := stsTotalPublished + 1;
        ELSE
            // Failure - track consecutive failures
            _signals[_signalIndex].nConsecFails := _signals[_signalIndex].nConsecFails + 1;
            _consecFailures := _consecFailures + 1;
            stsConsecFailures := _consecFailures;

            // Check fault threshold
            IF _consecFailures >= cfgMaxConsecFails THEN
                stsFaulted := TRUE;
                stsFaultCode := FAULT_PUBLISH;
                Run := FALSE;
                RETURN;
            END_IF
        END_IF
    END_IF

END_WHILE

// ─────────────────────────────────────────────────────────────────────
// TRANSACTION GROUP ENGINE - Publish grouped signals as JSON
// Each group collects all assigned signals and publishes a single
// JSON object: {"subtopic1":value1,"subtopic2":value2,...}
// ─────────────────────────────────────────────────────────────────────
FOR _txGroupIdx := 1 TO 3 DO

    // Get period and matching mode for this group
    CASE _txGroupIdx OF
        1:  _txGroupPeriod := cfgTxGroup1Period;
            _txGroupMode := E_MQTT_PublishMode.TRANSACTION_GROUP_1;
        2:  _txGroupPeriod := cfgTxGroup2Period;
            _txGroupMode := E_MQTT_PublishMode.TRANSACTION_GROUP_2;
        3:  _txGroupPeriod := cfgTxGroup3Period;
            _txGroupMode := E_MQTT_PublishMode.TRANSACTION_GROUP_3;
    END_CASE

    // Check if period has elapsed
    IF (_currentTime - _txGroupLastTime[_txGroupIdx]) < _txGroupPeriod THEN
        CONTINUE;
    END_IF

    // Build JSON payload
    MEMSET(ADR(_txPayload), 0, SIZEOF(_txPayload));
    _txLen := 0;
    AppendToPayload('{');
    _txFirst := TRUE;
    _txHasSignals := FALSE;

    FOR _i := 1 TO _signalCount DO
        IF NOT _signals[_i].bRegistered THEN
            CONTINUE;
        END_IF
        IF _signals[_i].ePublishMode <> _txGroupMode THEN
            CONTINUE;
        END_IF
        // Skip subscribe-only signals
        IF _signals[_i].eDirection = E_MQTT_Direction.SUBSCRIBE THEN
            CONTINUE;
        END_IF

        // Validate pointer
        IF NOT IsPointerValid(_signals[_i].pValue) THEN
            stsFaulted := TRUE;
            stsFaultCode := FAULT_POINTER_INVALID;
            Run := FALSE;
            RETURN;
        END_IF

        _txHasSignals := TRUE;

        // Add comma separator between entries
        IF NOT _txFirst THEN
            AppendToPayload(',');
        END_IF
        _txFirst := FALSE;

        // Add "key":value
        AppendToPayload('"');
        AppendToPayload(_signals[_i].sSubTopic);
        AppendToPayload('":');

        // Get value as string
        _currentValue := ValueToString(
            inpPValue := _signals[_i].pValue,
            inpType := _signals[_i].eType
        );

        // Quote string and time values for valid JSON
        IF _signals[_i].eType = E_MQTT_SignalType.TYPE_STRING
           OR _signals[_i].eType = E_MQTT_SignalType.TYPE_TIME THEN
            AppendToPayload('"');
            AppendToPayload(_currentValue);
            AppendToPayload('"');
        ELSE
            AppendToPayload(_currentValue);
        END_IF

        // Update last published value (for bidirectional re-publish suppression)
        _signals[_i].sLastPublished := _currentValue;
    END_FOR

    AppendToPayload('}');

    // Publish if there are signals in this group
    IF _txHasSignals THEN
        // Build full topic: cfgPublishBaseTopic/cfgTxGroupNTopic
        CASE _txGroupIdx OF
            1: _fullTopic := CONCAT(CONCAT(cfgPublishBaseTopic, '/'), cfgTxGroup1Topic);
            2: _fullTopic := CONCAT(CONCAT(cfgPublishBaseTopic, '/'), cfgTxGroup2Topic);
            3: _fullTopic := CONCAT(CONCAT(cfgPublishBaseTopic, '/'), cfgTxGroup3Topic);
        END_CASE

        _publishResult := mqttClient.Publish(
            sTopic := _fullTopic,
            pPayload := ADR(_txPayload),
            nPayloadSize := _txLen,
            eQoS := cfgPublishQoS,
            bRetain := cfgRetainPublish
        );

        IF _publishResult THEN
            _txGroupLastTime[_txGroupIdx] := _currentTime;
            _consecFailures := 0;
            stsTotalPublished := stsTotalPublished + 1;
        ELSE
            _consecFailures := _consecFailures + 1;
            stsConsecFailures := _consecFailures;
            IF _consecFailures >= cfgMaxConsecFails THEN
                stsFaulted := TRUE;
                stsFaultCode := FAULT_PUBLISH;
                Run := FALSE;
                RETURN;
            END_IF
        END_IF
    END_IF

END_FOR

// ─────────────────────────────────────────────────────────────────────
// SUBSCRIBE ENGINE - Process incoming messages from queue
// Supports raw payloads and JSON key extraction
// Multiple signals can share a topic (each extracts a different JSON key)
// ─────────────────────────────────────────────────────────────────────
WHILE mqttClient.fbMessageQueue.nQueuedMessages > 0 DO

    // Clear receive buffers
    MEMSET(ADR(_receivedTopic), 0, SIZEOF(_receivedTopic));
    MEMSET(ADR(_receivedPayload), 0, SIZEOF(_receivedPayload));

    // Dequeue next message
    IF NOT mqttClient.fbMessageQueue.Dequeue(fbMessage := mqttMessage) THEN
        EXIT;
    END_IF

    // Extract topic and payload
    mqttMessage.GetTopic(pTopic := ADR(_receivedTopic), nTopicSize := SIZEOF(_receivedTopic));
    mqttMessage.GetPayload(pPayload := ADR(_receivedPayload), nPayloadSize := SIZEOF(_receivedPayload), bSetNullTermination := TRUE);

    stsTotalReceived := stsTotalReceived + 1;

    // Parse JSON once per message if payload starts with '{'
    _jsonParsed := FALSE;
    IF LEN(_receivedPayload) > 0 AND_THEN _receivedPayload[0] = 16#7B THEN // 0x7B = '{'
        _jsonDoc := fbJsonParser.ParseDocument(_receivedPayload);
        _jsonRoot := fbJsonParser.GetDocumentRoot();
        _jsonParsed := fbJsonParser.IsObject(_jsonRoot);
    END_IF

    // Iterate ALL registered signals (multiple signals can share a topic)
    FOR _i := 1 TO _signalCount DO
        IF NOT _signals[_i].bRegistered THEN
            CONTINUE;
        END_IF

        // Check if direction allows subscribe/write
        IF _signals[_i].eDirection <> E_MQTT_Direction.SUBSCRIBE
           AND _signals[_i].eDirection <> E_MQTT_Direction.BIDIRECTIONAL THEN
            CONTINUE;
        END_IF

        // Match topic
        _fullTopic := CONCAT(CONCAT(cfgSubscribeBaseTopic, '/'), _signals[_i].sSubTopic);
        IF _fullTopic <> _receivedTopic THEN
            CONTINUE;
        END_IF

        // Validate pointer before writing
        IF NOT IsPointerValid(_signals[_i].pValue) THEN
            stsFaulted := TRUE;
            stsFaultCode := FAULT_POINTER_INVALID;
            Run := FALSE;
            RETURN;
        END_IF

        IF LEN(_signals[_i].sJsonKey) > 0 AND _jsonParsed THEN
            // JSON mode: extract specific key from parsed document
            _jsonValueStr := ExtractJsonValue(
                inpJsonKey := _signals[_i].sJsonKey,
                inpJsonParentKey := _signals[_i].sJsonParentKey
            );

            // Only write if key was found (non-empty result)
            IF LEN(_jsonValueStr) > 0 THEN
                StringToValue(
                    inpPayload := _jsonValueStr,
                    inpPValue := _signals[_i].pValue,
                    inpType := _signals[_i].eType
                );
                _signals[_i].sLastPublished := _jsonValueStr;
            END_IF

        ELSIF LEN(_signals[_i].sJsonKey) = 0 THEN
            // Raw mode: use entire payload as value (original behavior)
            StringToValue(
                inpPayload := _receivedPayload,
                inpPValue := _signals[_i].pValue,
                inpType := _signals[_i].eType
            );
            _signals[_i].sLastPublished := _receivedPayload;
        END_IF
        // If sJsonKey is set but JSON didn't parse, silently skip

    END_FOR

END_WHILE

Run := TRUE;
END_METHOD

// ═══════════════════════════════════════════════════════════════════════
// METHOD PRIVATE StringToValue
// Write string payload to pointer based on type
// Returns: TRUE if successful, FALSE if type not supported
// ═══════════════════════════════════════════════════════════════════════
METHOD PRIVATE StringToValue : BOOL
VAR_INPUT
    inpPayload  : STRING(255);
    inpPValue   : PVOID;
    inpType     : E_MQTT_SignalType;
END_VAR
VAR
    _pBool      : POINTER TO BOOL;
    _pByte      : POINTER TO BYTE;
    _pInt       : POINTER TO INT;
    _pDint      : POINTER TO DINT;
    _pReal      : POINTER TO REAL;
    _pLreal     : POINTER TO LREAL;
    _pString    : POINTER TO STRING(255);
    _pTime      : POINTER TO TIME;
    _upperPayload: STRING(255);
END_VAR
StringToValue := TRUE;

CASE inpType OF

    E_MQTT_SignalType.TYPE_BOOL:
        _pBool := inpPValue;
        _upperPayload := F_ToUCase(inpPayload);
        _pBool^ := (_upperPayload = 'TRUE') OR (_upperPayload = '1') OR (_upperPayload = 'ON');

    E_MQTT_SignalType.TYPE_BYTE:
        _pByte := inpPValue;
        _pByte^ := STRING_TO_BYTE(inpPayload);

    E_MQTT_SignalType.TYPE_INT:
        _pInt := inpPValue;
        _pInt^ := STRING_TO_INT(inpPayload);

    E_MQTT_SignalType.TYPE_DINT:
        _pDint := inpPValue;
        _pDint^ := STRING_TO_DINT(inpPayload);

    E_MQTT_SignalType.TYPE_REAL:
        _pReal := inpPValue;
        _pReal^ := STRING_TO_REAL(inpPayload);

    E_MQTT_SignalType.TYPE_LREAL:
        _pLreal := inpPValue;
        _pLreal^ := STRING_TO_LREAL(inpPayload);

    E_MQTT_SignalType.TYPE_STRING:
        _pString := inpPValue;
        _pString^ := inpPayload;

    E_MQTT_SignalType.TYPE_TIME:
        _pTime := inpPValue;
        _pTime^ := STRING_TO_TIME(inpPayload);

ELSE
    StringToValue := FALSE;
END_CASE
END_METHOD

// ═══════════════════════════════════════════════════════════════════════
// METHOD PRIVATE ValueToString
// Convert pointer value to string based on type
// ═══════════════════════════════════════════════════════════════════════
METHOD PRIVATE ValueToString : STRING(255)
VAR_INPUT
    inpPValue   : PVOID;
    inpType     : E_MQTT_SignalType;
END_VAR
VAR
    _pBool      : POINTER TO BOOL;
    _pByte      : POINTER TO BYTE;
    _pInt       : POINTER TO INT;
    _pDint      : POINTER TO DINT;
    _pReal      : POINTER TO REAL;
    _pLreal     : POINTER TO LREAL;
    _pString    : POINTER TO STRING(255);
    _pTime      : POINTER TO TIME;
END_VAR
CASE inpType OF

    E_MQTT_SignalType.TYPE_BOOL:
        _pBool := inpPValue;
        IF _pBool^ THEN
            ValueToString := 'true';
        ELSE
            ValueToString := 'false';
        END_IF

    E_MQTT_SignalType.TYPE_BYTE:
        _pByte := inpPValue;
        ValueToString := BYTE_TO_STRING(_pByte^);

    E_MQTT_SignalType.TYPE_INT:
        _pInt := inpPValue;
        ValueToString := INT_TO_STRING(_pInt^);

    E_MQTT_SignalType.TYPE_DINT:
        _pDint := inpPValue;
        ValueToString := DINT_TO_STRING(_pDint^);

    E_MQTT_SignalType.TYPE_REAL:
        _pReal := inpPValue;
        ValueToString := REAL_TO_STRING(_pReal^);

    E_MQTT_SignalType.TYPE_LREAL:
        _pLreal := inpPValue;
        ValueToString := LREAL_TO_STRING(_pLreal^);

    E_MQTT_SignalType.TYPE_STRING:
        _pString := inpPValue;
        ValueToString := _pString^;

    E_MQTT_SignalType.TYPE_TIME:
        _pTime := inpPValue;
        ValueToString := TIME_TO_STRING(_pTime^);

ELSE
    ValueToString := '';
END_CASE
END_METHOD

END_FUNCTION_BLOCK

// ---- POUs/FBs/fb_WriteDataToFile.TcPOU
FUNCTION_BLOCK  fb_WriteDataToFile
VAR_INPUT
    inpFilePath   : STRING(255);
    inpFileName   : STRING(255);
    data          : POINTER TO STRING;
	len			  : UDINT;
END_VAR
VAR_OUTPUT
    bBusy         : BOOL;
    bDone         : BOOL;
    bError        : BOOL;
    hrErrorId     : HRESULT;
END_VAR
VAR
    nState        : INT;
    trigExecute   : R_TRIG;
    bExecute      : BOOL;
    sFullFilePath : STRING(255);
    hFile         : UINT := 0;
    fbFileOpen    : FB_FileOpen;
    fbFileWrite   : FB_FileWrite;
    fbFileClose   : FB_FileClose;
END_VAR

trigExecute(CLK:=bExecute);

IF NOT bExecute THEN
    bDone := FALSE;
END_IF;

CASE nState OF
    0:
        bBusy := FALSE;
        bError := FALSE;
        hrErrorId := 0;
		

        IF trigExecute.Q THEN
            bBusy := TRUE;
            bDone := FALSE;
            bError := FALSE;
            sFullFilePath := '';
            nState := 10;
        END_IF;

    10:
        sFullFilePath := CONCAT(inpFilePath, '\');
		sFullFilePath := CONCAT(sFullFilePath, inpFileName);
        fbFileOpen(
            bExecute    := TRUE,
            sNetId      := '',
            sPathName   := sFullFilePath,
            nMode       := FOPEN_MODEWRITE,
            ePath       := PATH_GENERIC,
            tTimeout    := T#5S
        );
        nState := 20;

    20:
        fbFileOpen(bExecute := FALSE);

        IF NOT fbFileOpen.bBusy THEN
            IF fbFileOpen.bError THEN
                hrErrorId := TO_DINT(fbFileOpen.nErrId);
                nState := 99;
            ELSE
                hFile := fbFileOpen.hFile;
                nState := 30;
            END_IF;
        END_IF;

    30:
        fbFileWrite(
            bExecute    := TRUE,
            sNetId      := '',
            hFile       := hFile,
            pWriteBuff  := data,
            cbWriteLen  := len,
            tTimeout    := T#5S
        );
        nState := 40;

    40:
        fbFileWrite(bExecute := FALSE);

        IF NOT fbFileWrite.bBusy THEN
            IF fbFileWrite.bError THEN
                hrErrorId := TO_DINT(fbFileWrite.nErrId);
                nState := 80;
            ELSE
                nState := 50;
            END_IF;
        END_IF;

    50:
        fbFileClose(
            bExecute    := TRUE,
            sNetId      := '',
            hFile       := hFile,
            tTimeout    := T#5S
        );
        nState := 60;

    60:
        fbFileClose(bExecute := FALSE);

        IF NOT fbFileClose.bBusy THEN
            IF fbFileClose.bError THEN
                hrErrorId := TO_DINT(fbFileClose.nErrId);
                nState := 99;
            ELSE
                bDone := TRUE;
                bExecute := FALSE;
                nState := 0;
            END_IF;
        END_IF;

    80:
        fbFileClose(bExecute := TRUE, hFile := hFile);
        IF NOT fbFileClose.bBusy THEN
             nState := 99;
        END_IF;

    99:
        bError := TRUE;
        bBusy := FALSE;
        bExecute := FALSE;

        fbFileOpen(bExecute := FALSE);
        fbFileWrite(bExecute := FALSE);
        fbFileClose(bExecute := FALSE);

        IF NOT trigExecute.Q THEN
            nState := 0;
        END_IF;

END_CASE;

METHOD write : BOOL
VAR_INPUT
END_VAR
IF nState = 0 THEN
    bExecute := TRUE;
    Write := TRUE;
ELSE
    Write := FALSE;
END_IF;
END_METHOD

END_FUNCTION_BLOCK

// ---- POUs/FBs/Devices/fb_Dev_Actuator.TcPOU
FUNCTION_BLOCK fb_Dev_Actuator EXTENDS abs_fb_Device
VAR_INPUT
	IO_Input_Feedback : BOOL;
END_VAR

VAR_IN_OUT
	IO_Output_Actuate : BOOL;
END_VAR

VAR
	HMI						: ST_Actuator_HMI_Interface;
	_setActuate 			: BOOL;
	_retractOnFault			: BOOL;
	_hasFeedback			: BOOL;
	_faultH_onDelay			: TON;
	_faultH_offDelay		: TON;
	_faultH_OnDelay_Trigger	: BOOL;
	_faultH_OffDelay_Trigger: BOOL;
	_onDelay_time			: TIME;
	_offDelay_time			: TIME;
	_InvFeedback			: BOOL;
	_actuatorFeedback		: BOOL;
	_maintainAutoState		: BOOL;
	_disableHMIControl		: BOOL;
END_VAR

VAR_OUTPUT
	stsActuated : BOOL;

END_VAR

DeviceLogic();
Interlock.name := _DeviceName;
Interlock(inpConfig := _dataInterlock);

// Flip feedback if cofigured for inverted feedback
IF _InvFeedback THEN
	IF IO_Input_Feedback THEN
		_actuatorFeedback := FALSE;
	ELSE
		_actuatorFeedback :=TRUE;
	END_IF
ELSE
	IF IO_Input_Feedback THEN
		_actuatorFeedback :=TRUE;
	ELSE
		_actuatorFeedback :=FALSE;
	END_IF
END_IF

// If no IO based feedback, set actuation state for feedback
IF _hasFeedback THEN
	stsActuated := _actuatorFeedback;
ELSE
	stsActuated := _setActuate;
END_IF

// Check for timeouts
FaultHandler(_actuatorFeedback);

// Control via HMI if in manual
// cmdActuate an cmdRetract methods only work in Auto, unless
// device is configured for no manual control
IF NOT _disableHMIControl THEN
	IF NOT _inAuto THEN 
		IF HMI.ocmdActuate THEN
			cmdActuate();
		ELSE
			cmdRetract();
		END_IF
	ELSE
		// if property set, change the HMI actuatoion toggle state so that
		// transition from auto to manual does not change the state
		// otherwise upon transition HMI will change state to whatever it was in manual last
		IF _maintainAutoState THEN
			HMI.ocmdActuate := _setActuate;
		END_IF
	END_IF
END_IF
// Configure retract on feedback
IF stsFaulted AND _retractOnFault THEN
	HMI.ocmdActuate := 0;
	_setActuate		:= 0;
END_IF

// Log state changes
IF _setActuate THEN
	IO_output_actuate :=TRUE;
	sendLog('Actuating ON',1);
ELSE
	IO_output_actuate :=FALSE;
	sendLog('Actuating OFF',1);
END_IF

HMI.HMIbaseDevice := HMIbaseDevice;
HMI.stsActuated   := stsActuated;
HMI.setActuate    := _setActuate;

PROPERTY cfgDeviceName : string
GET
cfgDeviceName := _DeviceName;
END_GET
SET
_DeviceName := cfgDeviceName;
END_SET
END_PROPERTY

PROPERTY cfgDisableHMIControl : BOOL
GET
cfgDisableHMIControl := _disableHMIControl;
END_GET
SET
_disableHMIControl := cfgDisableHMIControl;
END_SET
END_PROPERTY

PROPERTY cfgHasFeedback : BOOL
GET
cfgHasFeedback := _hasFeedback;
END_GET
SET
_hasFeedback	:= cfgHasFeedback;
END_SET
END_PROPERTY

PROPERTY PUBLIC cfgInvFeedback : Bool
GET
cfgInvFeedback := _InvFeedback;
END_GET
SET
_InvFeedback := cfgInvFeedback;
END_SET
END_PROPERTY

PROPERTY cfgMaintainAutoState : BOOL
GET
cfgMaintainAutoState	:= _maintainAutoState;
END_GET
SET
_maintainAutoState := cfgMaintainAutoState;
END_SET
END_PROPERTY

PROPERTY cfgOffDelay : TIME
GET
cfgOffDelay := _offDelay_time;
END_GET
SET
_offDelay_time := cfgOffDelay;
END_SET
END_PROPERTY

PROPERTY PUBLIC cfgOnDelay : Time
GET
cfgOnDelay := _onDelay_time;
END_GET
SET
_OnDelay_time := cfgOnDelay;
END_SET
END_PROPERTY

PROPERTY cfgRetractOnFault : bool
GET
cfgRetractOnFault := _retractOnFault;
END_GET
SET
_retractOnFault := cfgRetractOnFault;
END_SET
END_PROPERTY

METHOD PUBLIC cmdActuate : BOOL
VAR_INPUT
	
END_VAR
IF Interlock.outInterlockOK AND NOT stsFaulted THEN
	_setActuate :=TRUE;
END_IF
END_METHOD

METHOD cmdReset : BOOL
IF stsFaulted THEN
	setFault(0,'');
END_IF
END_METHOD

METHOD PUBLIC cmdRetract : BOOL
VAR_INPUT
END_VAR
// Retracting (de-energising) is always allowed. It used to require the interlock to be met,
// so an actuator whose interlock dropped could not be switched off, by the operator or by code,
// unless cfgRetractOnFault happened to be set.
_setActuate := FALSE;
END_METHOD

METHOD PRIVATE FaultHandler : BOOL
VAR_INPUT
	inpFeedback : BOOL; 
	
END_VAR
//if setActuate, set timer. If timer done and no feedback, then fault
IF (_onDelay_Time <> T#0S) AND _hasfeedback THEN
	_faultH_onDelay(IN:=_faultH_OnDelay_Trigger,PT:=_onDelay_time);
	IF (NOT stsFaulted) AND _setActuate THEN
		_faultH_OnDelay_Trigger := TRUE;
		IF _faultH_onDelay.Q AND NOT _actuatorFeedback THEN
			setFault(1,'actuator feedback missing.');
		END_IF
	ELSE
		_faultH_OnDelay_Trigger := FALSE;
	END_IF
END_IF

IF (_offDelay_Time <> T#0S) AND _hasfeedback THEN
	_faultH_offDelay(IN:=_faultH_OffDelay_Trigger,PT:=_offDelay_time);
	IF (NOT stsFaulted) AND NOT(_setActuate) THEN
		_faultH_OffDelay_Trigger := TRUE;
		IF _faultH_offDelay.Q AND _actuatorFeedback THEN
			setFault(1,'Feedback present when not actuated.');
		END_IF
	ELSE
		_faultH_OffDelay_Trigger := FALSE;
	END_IF
END_IF


//IF _actuatorFeedback AND NOT(_setActuate) and _hasFeedback THEN
//	setFault(1,'Feedback present when not actuated');
//END_IF

//if not actuated but feedback is in, actuator is stuck closed
//+TODO

//If enabled and cmdActuated and lost interlock, then fault
IF NOT stsFaulted AND _setActuate THEN
	IF NOT interlock.outInterlockOK THEN
		setFault(1,CONCAT('I_NOK - ',Interlock.stsFirstOut));
	END_IF
END_IF
END_METHOD

//FB_Init is always available implicitly and it is used primarily for initialization.
//The return value is not evaluated. For a specific influence, you can also declare the
//methods explicitly and provide additional code there with the standard initialization
//code. You can evaluate the return value.
METHOD FB_Init: BOOL
VAR_INPUT
    bInitRetains: BOOL; // TRUE: the retain variables are initialized (reset warm / reset cold)
    bInCopyCode: BOOL;  // TRUE: the instance will be copied to the copy code afterward (online change)
	
	cfgDeviceName 		: STRING;
	cfgEnable 			: BOOL;
	cfgInitEventClass	: BOOL;
	cfgOnDelay 			: TIME;
	cfgOffDelay			: TIME;
	cfgRetractOnFault 	: BOOL;
	cfgInvFeedback		: BOOL; 
	cfgHasFeedback		: BOOL;

END_VAR
THIS^.cfgDeviceName 		:= 		cfgDeviceName; 
THIS^.cfgEnable				:=		cfgEnable;
THIS^.cfgInitEventClass		:= 		cfgInitEventClass;		
THIS^.cfgOnDelay 			:= 		cfgOnDelay; 
THIS^.cfgOffDelay			:=		cfgOffDelay;			
THIS^.cfgRetractOnFault		:=      cfgRetractOnFault;
THIS^.cfgInvFeedback		:=		cfgInvFeedback;
THIS^.cfgHasFeedback		:=		cfgHasFeedback;
END_METHOD

END_FUNCTION_BLOCK

// ---- POUs/FBs/Devices/fb_Dev_XPendant.TcPOU
(*
    fb_Dev_XPendant — Xbox-controller pendant endpoint.

    The lhmi sidecar app `xpendant` (lhmi-core apps/xpendant) reads a USB Xbox
    controller on the IPC and writes its state into the public Pad member over local ADS — the
    FB instance path is passed to that service as an argument, and the member
    names of ST_XPendant_In are the write contract (<instance>.Pad.<member>). This FB only OUTPUTS what
    the controller is doing; wiring those outputs to motion is machine logic, outside this FB.

    Analog outputs = DIRECTION + SPEED (jog-ready). Each stick axis and each trigger
    is broken into an ST_XPendant_Axis { Value, Pos, Neg, Throttle }:
      Pos/Neg = which way it's pushed past cfgActivateThreshold (jog direction);
        sticks are bidirectional (Pos = up/right, Neg = down/left), triggers are
        one-sided (Pos = pulled, Neg always FALSE).
      Throttle = 0..100 % magnitude ("how far") = a custom speed override; 0 unless
        Pos or Neg is set.
    So "left analog up @ 70 %" is stsLeftStickY.Pos = TRUE, stsLeftStickY.Throttle = 70.

    Liveness contract: the service bumps Pad.Watchdog every ~500 ms and holds
    Pad.Connected while a controller is present. stsFeedAlive drops when the
    watchdog stops changing for cfgFeedTimeout (default T#1S500MS = 3 missed
    beats); ALL outputs are zeroed unless stsConnected. Consumers must still
    apply their own gating (e.g. a held dead-man on an axis) — this FB is an
    input device, never a safety path.

    Supervision: inpActive (machine logic) declares when the pendant is EXPECTED —
    unplugged is the normal state for a teach pendant, so absence is only
    warning-worthy while inpActive is TRUE (the IPC service reads the mirror
    HMI.Status.stsInService and drives the HMI warning). inpActive does not gate outputs.

    Usage:
        XPendant : fb_Dev_XPendant(cfgDeviceName := 'XPendant', cfgEnable := TRUE,
                                   cfgInitEventClass := TRUE, cfgFeedTimeout := T#1S500MS);
        XPendant(inpAuto := Machine.stsInAuto, inpReset := Machine.cmdReset,
                 inpInterlockBypass := FALSE, faultMonitor := ADR(FaultMonitor),
                 inpActive := <machine logic: pendant operation selected>);
        // jog an axis from the left stick's Y (up/down), speed from how far it's pushed:
        Axis1(inpPendantJogPos := XPendant.stsLeftStickY.Pos,
              inpPendantJogNeg := XPendant.stsLeftStickY.Neg,
              inpPendantJogVelo := cfgJogMax * XPendant.stsLeftStickY.Throttle / 100.0);
*)
FUNCTION_BLOCK fb_Dev_XPendant EXTENDS abs_fb_Device
VAR_INPUT
    // SUPERVISION flag, driven by machine logic: TRUE = the pendant is expected /
    // in service right now (e.g. manual mode + pendant operation selected). A teach
    // pendant is exceptional equipment — unplugged is the NORMAL state — so while
    // FALSE (the default) nothing anywhere complains about an absent controller;
    // while TRUE, absence is warning-worthy (the IPC service reads the mirror
    // HMI.Status.stsInService and raises the HMI warning). Does NOT gate the pad
    // outputs: a plugged, live controller always passes through — consumers keep
    // their own gating.
    inpActive : BOOL;
END_VAR

VAR_OUTPUT
    stsConnected : BOOL;    // controller present AND feed alive AND device enabled
    stsFeedAlive : BOOL;    // service watchdog fresh (Pad.Watchdog changed within cfgFeedTimeout)
    stsActive    : BOOL;    // inpActive AND stsConnected — "pendant in service and usable now"

    // Gated pad state — all FALSE / 0.0 while NOT stsConnected:
    stsBtnA      : BOOL;
    stsBtnB      : BOOL;
    stsBtnX      : BOOL;
    stsBtnY      : BOOL;
    stsBumpL     : BOOL;
    stsBumpR     : BOOL;
    stsStart     : BOOL;
    stsBack      : BOOL;
    stsThumbL    : BOOL;    // left-stick click (L3)
    stsThumbR    : BOOL;    // right-stick click (R3)
    stsDpadUp    : BOOL;
    stsDpadDown  : BOOL;
    stsDpadLeft  : BOOL;
    stsDpadRight : BOOL;

    // Analog controls as DIRECTION + SPEED pairs (ST_XPendant_Axis). Sticks are
    // bidirectional (Pos = up/right, Neg = down/left); triggers are one-sided (Pos
    // = pulled, Neg always FALSE). Throttle = 0..100 %. See the header for wiring.
    stsLeftStickX  : ST_XPendant_Axis;
    stsLeftStickY  : ST_XPendant_Axis;
    stsRightStickX : ST_XPendant_Axis;
    stsRightStickY : ST_XPendant_Axis;
    stsTriggerL    : ST_XPendant_Axis;   // LT
    stsTriggerR    : ST_XPendant_Axis;   // RT
END_VAR

VAR
    // Written over ADS by the xpendant IPC service (raw external mirror — never
    // drive from PLC logic). A plain VAR on purpose: FB VAR_INPUT members are not
    // reliably in the ADS symbol download (the cfgUnit/1808 lesson), while public
    // VAR members — the same surface as HMI below — are.
    Pad          : ST_XPendant_In;

    HMI          : ST_XPendant_HMI_Interface;   // Public HMI interface — bind <instance>.HMI
    _wdLast      : UINT;                        // last seen watchdog count
    _wdStale     : TON;                         // runs while the watchdog is UNCHANGED
    _feedTimeout : TIME := T#1S500MS;           // see cfgFeedTimeout
    _activateThreshold : LREAL := 0.05;         // deflection (fraction) before Pos/Neg engage — see cfgActivateThreshold
END_VAR

// ── 1. Base device logic (init, interlock, faults, reset, HMIbaseDevice) ──
DeviceLogic();

// ── 2. Feed liveness. The service bumps Pad.Watchdog every ~500 ms; the TON
//       runs while the count is UNCHANGED, so expiry = the feed went stale/dead
//       (same time-since-last-good-data idiom as the Modbus driver). ──
_wdStale(IN := (Pad.Watchdog = _wdLast), PT := _feedTimeout);
stsFeedAlive := NOT _wdStale.Q;
IF Pad.Watchdog <> _wdLast THEN
    _wdLast := Pad.Watchdog;
END_IF

stsConnected := Pad.Connected AND stsFeedAlive AND _enabled;
stsActive    := inpActive AND stsConnected;

// ── 3a. Buttons: gated pass-through — outputs mirror the pad ONLY while connected ──
IF stsConnected THEN
    stsBtnA      := Pad.BtnA;
    stsBtnB      := Pad.BtnB;
    stsBtnX      := Pad.BtnX;
    stsBtnY      := Pad.BtnY;
    stsBumpL     := Pad.BumpL;
    stsBumpR     := Pad.BumpR;
    stsStart     := Pad.Start;
    stsBack      := Pad.Back;
    stsThumbL    := Pad.ThumbL;
    stsThumbR    := Pad.ThumbR;
    stsDpadUp    := Pad.DpadUp;
    stsDpadDown  := Pad.DpadDown;
    stsDpadLeft  := Pad.DpadLeft;
    stsDpadRight := Pad.DpadRight;
ELSE
    stsBtnA      := FALSE;
    stsBtnB      := FALSE;
    stsBtnX      := FALSE;
    stsBtnY      := FALSE;
    stsBumpL     := FALSE;
    stsBumpR     := FALSE;
    stsStart     := FALSE;
    stsBack      := FALSE;
    stsThumbL    := FALSE;
    stsThumbR    := FALSE;
    stsDpadUp    := FALSE;
    stsDpadDown  := FALSE;
    stsDpadLeft  := FALSE;
    stsDpadRight := FALSE;
END_IF

// ── 3b. Analogs -> direction trigger + 0..100 % throttle (deriveAxis). Feed the
//        gated raw value: 0.0 when not connected yields a fully-zeroed axis. ──
IF stsConnected THEN
    stsLeftStickX  := deriveAxis(Pad.StickLX, TRUE);
    stsLeftStickY  := deriveAxis(Pad.StickLY, TRUE);
    stsRightStickX := deriveAxis(Pad.StickRX, TRUE);
    stsRightStickY := deriveAxis(Pad.StickRY, TRUE);
    stsTriggerL    := deriveAxis(Pad.TrigL, FALSE);
    stsTriggerR    := deriveAxis(Pad.TrigR, FALSE);
ELSE
    stsLeftStickX  := deriveAxis(0.0, TRUE);
    stsLeftStickY  := deriveAxis(0.0, TRUE);
    stsRightStickX := deriveAxis(0.0, TRUE);
    stsRightStickY := deriveAxis(0.0, TRUE);
    stsTriggerL    := deriveAxis(0.0, FALSE);
    stsTriggerR    := deriveAxis(0.0, FALSE);
END_IF

// ── 4. Publish to HMI ──
HMI.HMIbaseDevice        := HMIbaseDevice;
HMI.Status.stsConnected  := stsConnected;
HMI.Status.stsFeedAlive  := stsFeedAlive;
HMI.Status.stsActive     := stsActive;
HMI.Status.stsInService  := inpActive;   // supervision mirror — the IPC service READS this
HMI.Status.stsBtnA       := stsBtnA;
HMI.Status.stsBtnB       := stsBtnB;
HMI.Status.stsBtnX       := stsBtnX;
HMI.Status.stsBtnY       := stsBtnY;
HMI.Status.stsBumpL      := stsBumpL;
HMI.Status.stsBumpR      := stsBumpR;
HMI.Status.stsStart      := stsStart;
HMI.Status.stsBack       := stsBack;
HMI.Status.stsThumbL     := stsThumbL;
HMI.Status.stsThumbR     := stsThumbR;
HMI.Status.stsDpadUp     := stsDpadUp;
HMI.Status.stsDpadDown   := stsDpadDown;
HMI.Status.stsDpadLeft   := stsDpadLeft;
HMI.Status.stsDpadRight  := stsDpadRight;
HMI.Status.stsLeftStickX  := stsLeftStickX;
HMI.Status.stsLeftStickY  := stsLeftStickY;
HMI.Status.stsRightStickX := stsRightStickX;
HMI.Status.stsRightStickY := stsRightStickY;
HMI.Status.stsTriggerL    := stsTriggerL;
HMI.Status.stsTriggerR    := stsTriggerR;

// Watchdog staleness threshold. Service beats ~500 ms; default 1.5 s = 3 missed beats.
PROPERTY cfgFeedTimeout : TIME
GET
cfgFeedTimeout := _feedTimeout;
END_GET
SET
IF cfgFeedTimeout > T#0MS THEN
    _feedTimeout := cfgFeedTimeout;
END_IF
END_SET
END_PROPERTY

// Deflection (0..1 fraction) a stick/trigger must exceed before Pos/Neg engage and
// Throttle leaves 0. The service already applies XInput dead zones and rescales to
// 0..1, so this is a small extra jog-arming margin (default 0.05 = 5 %). Property
// only (no FB_Init param) so it never disturbs an existing instance declaration.
PROPERTY cfgActivateThreshold : LREAL
GET
cfgActivateThreshold := _activateThreshold;
END_GET
SET
IF cfgActivateThreshold >= 0.0 AND cfgActivateThreshold < 1.0 THEN
    _activateThreshold := cfgActivateThreshold;
END_IF
END_SET
END_PROPERTY

// Break one raw analog value into a DIRECTION trigger + a 0..100 % speed throttle.
// allowNeg = TRUE for sticks (bidirectional), FALSE for triggers (+ only).
METHOD PRIVATE deriveAxis : ST_XPendant_Axis
VAR_INPUT
    value    : LREAL;
    allowNeg : BOOL;
END_VAR
deriveAxis.Value := value;
deriveAxis.Pos   := value > _activateThreshold;
deriveAxis.Neg   := allowNeg AND (value < (-1.0 * _activateThreshold));
IF deriveAxis.Pos OR deriveAxis.Neg THEN
    deriveAxis.Throttle := LIMIT(0.0, ABS(value) * 100.0, 100.0);
ELSE
    deriveAxis.Throttle := 0.0;
END_IF
END_METHOD

METHOD FB_Init : BOOL
VAR_INPUT
    bInitRetains      : BOOL; // TRUE: the retain variables are initialized (reset warm / reset cold)
    bInCopyCode       : BOOL; // TRUE: the instance will be copied to the copy code afterward (online change)
    cfgDeviceName     : STRING;
    cfgEnable         : BOOL;
    cfgInitEventClass : BOOL;
    cfgFeedTimeout    : TIME;
END_VAR
THIS^.cfgDeviceName     := cfgDeviceName;
THIS^.cfgEnable         := cfgEnable;
THIS^.cfgInitEventClass := cfgInitEventClass;
IF cfgFeedTimeout > T#0MS THEN
    _feedTimeout := cfgFeedTimeout;
END_IF
END_METHOD

// Standard accessor: expose the HMI struct to callers (house pattern, see fb_Axis).
METHOD PUBLIC getHMIdata : ST_XPendant_HMI_Interface
VAR_INPUT
END_VAR
getHMIdata := HMI;
END_METHOD

END_FUNCTION_BLOCK

// ---- POUs/FBs/Devices/fb_Dev_AnalogSensor.TcPOU
FUNCTION_BLOCK fb_Dev_AnalogSensor EXTENDS abs_fb_Device
VAR_INPUT
	inpRawIOChannel			: DINT;
	inpScaledIOChannel		: LREAL;
	inpChannelDiag			: ST_AnalogSensor_Diag; //IO channel diagnostics
	cfgScalingNeeded		: BOOL;					// Set to False if scaled in IO
	cfgChannelMinInt		: DINT;					//Min INT IO channel value
	cfgChannelMaxInt		: DINT;					//Max INT IO channel value
	cfgSensorMin			: LREAL;  				//Min Sensor value (0V, 4mA etc)
	cfgSensorMax			: LREAL;  				//Max Sensor value (10V, 20mA etc)
	cfgEngUnitMin			: LREAL;  				//Min span of instrument
	cfgEngUnitMax			: LREAL;  				//Max span of instrument

END_VAR
VAR_OUTPUT
	stsSensorRawSignal		: LREAL;
	stsEngValue				: LREAL;
END_VAR
VAR
	_sensorRawSignal		: LREAL;
	_engValue				: LREAL;
	_alarmEnable	: BOOL;
	_alarmL			: LREAL;
	_alarmLL		: LREAL;
	_alarmH			: LREAL;
	_alarmHH		: LREAL;
	_calOffset		: LREAL;
	_calGain		: LREAL := 1.0;	// 1 = no gain correction (0 would zero every reading)
	_engUnit		: STRING;
	_alarmDebounce  : ARRAY[1..4] OF TON;
	_alarmCooldown	: ARRAY[1..4] OF BOOL;
END_VAR

VAR PERSISTENT
	HMI	: ST_AnalogSensor_HMI_Interface;
END_VAR

DeviceLogic();

scaleInput();

FaultHandler();

setHMI();

stsSensorRawSignal	:= _sensorRawSignal;
stsEngValue			:= _engValue;

PROPERTY cfgAlarmEnable : BOOL
GET
cfgAlarmEnable := _alarmEnable;
END_GET
SET
_alarmEnable := cfgAlarmEnable;
END_SET
END_PROPERTY

